(* IEC 61131-3 sources: daoli-st-library/DL_Process (part 32) *)

(* ---- FB_DL_ElectrolyzerStackPurgeSeq.st ---- *)
//==============================================================================
// 功能块：FB_DL_ElectrolyzerStackPurgeSeq ｜ 中文名称：电解槽氮气吹扫与升压序（复杂度 C4）
// 所属子库：DL_Process ｜ 版本 VERSION: v1.0.0 ｜ 兼容：CODESYS V3.5+ / TwinCAT 3 / 汇川 InoProShop
// 功能描述：电解槽停机检修后的投运前置序——低压氮气保压检漏 → N2 置换吹扫（按置换
//           倍数 n = ln(C0/C1) 算所需体积）→ O2 校验 → 升压至运行压力 → 就绪放行
//           （H2 侧仅在就绪相且 O2 合格时才允许打开）→ 泄压走 eVent 单向。泄漏率超
//           限、吹扫/升压超时、O2 不合格一律不放行并锁存故障。
// 开源溯源 (Origin)：道莅原创实现（参考 ISO 22734 水电解制氢系统与 GB/T 19774 水
//           电解制氢系统技术要求 分类与参数域，许可证=MIT，借鉴点=「惰性气体置换至
//           爆炸下限以下再投氢」的置换倍数判据与硬互锁序）
// 单位表：O2[%] / 压力[bar] / 流量[Nm³/h] / 体积[Nm³] / 泄漏率[bar/min] / 时间[ms]
// 置换倍数公式（本件核心判据，单位与推导写清）：
//   n = ln(C0 / C1)；C0 = 空气 O2 体积分数 20.9 [%]，C1 = 目标 O2 阈值 1.0 [%]
//   → n = ln(20.9 / 1.0) ≈ 3.04 [倍]，即需通入约 3.04 倍栈容积的 N2。
//   累计 N2 体积 [Nm³] = Σ (fN2FlowNm3h ÷ 3600 × Δt[s])，Δt 取 DL_ELZ_DT_S 假定任务
//   周期 10 ms；置换倍数出口 = 累计体积 ÷ 栈容积 [倍]。除零由段 3/段 4 双侧闸拦。
// 错误码表（Process 段 0005，故障窗口 3F01~3F09，信息窗口 3F81/3F82）：
//   16#0005_3F01 故障级：组态非法（栈容积/目标压/泄漏限/时间量 <= 0 或 O2 阈值域外）
//   16#0005_3F02 故障级：实时量入口非有限（O2 / 压力 / 流量 NaN 或 Inf），拒算
//   16#0005_3F03 故障级：检修保压检漏超限（泄漏率 > fLeakLimitBarPerMin，不放行）
//   16#0005_3F04 故障级：吹扫超时（tPurgeMaxTime 内置换倍数未达 n）
//   16#0005_3F05 故障级：O2 校验失败（校验窗内 O2 未降至阈值以下）
//   16#0005_3F06 故障级：升压超时（预充压或正式升压未达目标压）
//   16#0005_3F07 故障级：投运前保压检漏超限（就绪相保压窗内泄漏率超限，不放行）
//   16#0005_3F08 故障级兜底：状态机落 ELSE 非法态，全输出断
//   16#0005_3F09 故障级：H2 硬互锁违反（就绪相 O2 回升超阈值，立即关 H2 并锁存）
//   16#0005_3F81 信息级：置换倍数达标（置换完成拍，不置 bError）
//   16#0005_3F82 信息级：系统就绪放行（进入 eReady 拍，不置 bError）
//           故障级码全部锁存回放（R187），唯一清除路径 = bReset 上升沿。
// 状态机：E_DL_ElyzPurgeState（八态：eIdle=0 / eLeakTest=10 / ePurge=20 / eVerifyO2=30 /
//           ePressurize=40 / eReady=50 / eVent=60 / eFault=99）。eVent 为单向泄压相，
//           迁出唯一目标 = eIdle，不得返回 eReady（防止带氢泄压后直接投运）。
// 边界行为：① H2 侧硬互锁三重闸：相位必须是 eReady、O2 <= 阈值、无任何故障锁存；段 8
//           的 CASE ELSE 与出口断言各断一次（双保险）；② O2 未达标绝不进 eReady，故
//           不可能放 H2；③ 泄漏率判据只用「>」单侧直比（泄漏率本身是统计量，不设容差
//           死区，避免漏判）；④ 八态 CASE 每态显式 + ELSE 兜底 → 3F08 全断；⑤ 中止在
//           任何运行相都只迁入 eVent（单向泄压），不走「原地停机」路径。
// 语义假设：① fO2Pct 为栈内气相 O2 体积分数，单位 %；② fLeakDropBarPerMin 由上层
//           压降速率仪表或本库泄漏率估算件提供（本件不重复实现估算）；③ N2 流量为
//           标况体积流量，压力对体积的修正由上层完成；④ 栈容积含管路死体积。
// 依赖纪律：仅 Standard.library（TON / R_TRIG / LN）；零 GVL、零 VAR_EXTERNAL、零物
//           理地址直连，业务侧只经引脚注入。
// 修订历史：v1.0.0 2026-11-25 R88 首版（无人值守批次 · 复杂件 C4 · 序号 3）
//==============================================================================

(*------------------------------------------------------------------------------
 * 枚举: E_DL_ElyzPurgeState（归属本功能块，同文件发布，全库唯一定义）
 * 含义: 吹扫升压相位，与段 7 状态机、段 8 输出置位一一对应。
 *-----------------------------------------------------------------------------*)
TYPE E_DL_ElyzPurgeState :
(
    eIdle       := 0,  // 空闲：等启动沿 / Idle, awaiting the start edge
    eLeakTest   := 10, // 检修检漏：低压氮气保压测泄漏率 / Leak test at low nitrogen pressure
    ePurge      := 20, // 吹扫：N2 置换至置换倍数达标 / Purge until the exchange ratio is reached
    eVerifyO2   := 30, // O2 校验：静置取样，O2 须稳定在阈值下 / O2 verification with a stable sample
    ePressurize := 40, // 升压：N2 升至运行压力 / Pressurise to the operating pressure
    eReady      := 50, // 就绪：放行相，H2 侧唯一允许投运的相位 / Ready, the only phase allowing H2
    eVent       := 60, // 泄压：单向排空至常压 / Vent, one-way depressurisation
    eFault      := 99  // 故障：泄漏/超时/O2/互锁/非法态 / Fault, leak, timeout, O2, interlock or illegal state
);
END_TYPE

FUNCTION_BLOCK FB_DL_ElectrolyzerStackPurgeSeq
VAR_INPUT
    xEnable             : BOOL;   // 使能，FALSE 期间按中止处理（转泄压） [—] / Enable, a drop aborts into venting
    xStart              : BOOL;   // 启动请求，上升沿生效 [—] / Start request, rising edge effective
    xAbort              : BOOL;   // 中止请求，任意拍生效，转 eVent 单向泄压 [—] / Abort request, moves to one-way venting
    xReset              : BOOL;   // 故障复位，上升沿清全部锁存 [—] / Fault reset, rising edge clears all latches
    fO2Pct              : LREAL;  // 栈内气相 O2 体积分数 [%] / Gas-phase O2 volume fraction [%]
    fStackPressBar      : LREAL;  // 栈内实际压力 [bar] / Actual stack pressure [bar]
    fTargetPressBar     : LREAL;  // 运行目标压力 [bar]，须 > 0 / Operating target pressure [bar]
    fN2FlowNm3h         : LREAL;  // 氮气标况流量 [Nm³/h] / Nitrogen normal-volume flow [Nm3/h]
    fStackVolM3         : LREAL;  // 栈与管路总容积 [Nm³]，须 > 0 / Total stack and piping volume [Nm3]
    fLeakDropBarPerMin  : LREAL;  // 实测压力下降速率 [bar/min] / Measured pressure decay rate [bar/min]
    fLeakLimitBarPerMin : LREAL;  // 允许泄漏率上限 [bar/min]，须 > 0 / Allowed leak rate ceiling [bar/min]
    tPurgeMaxTime       : TIME;   // 吹扫最长允许时间 [ms] / Maximum purge time [ms]
    tHoldTime           : TIME;   // 保压/取样稳定窗 [ms] / Hold and sampling window [ms]
    tPressTimeout       : TIME;   // 升压与预充压超时 [ms] / Pressurisation timeout [ms]
END_VAR
VAR_OUTPUT
    xN2ValveCmd         : BOOL;   // 氮气进气阀命令 [—] / Nitrogen inlet valve command
    xVentValveCmd       : BOOL;   // 排放阀命令（吹扫出口与泄压共用） [—] / Vent valve command
    xH2ValveCmd         : BOOL;   // 氢气侧阀命令（仅就绪相且 O2 合格才允许） [—] / H2 valve, ready phase and O2 proven only
    bRunning            : BOOL;   // 顺控运行中（非空闲非就绪非故障非泄压） [—] / Sequencing active
    bDone               : BOOL;   // 就绪放行电平（eReady 相） [—] / Ready-released level in the eReady phase
    bError              : BOOL;   // 故障级标志，仅故障级码置位 [—] / Fault-class flag, fault-level codes only
    nErrCode            : UDINT;  // 错误码，0 = 无错 [—] / Error code, 0 = none
    fPurgeVolRatio      : LREAL;  // 置换倍数出口 [倍] = 累计 N2 体积 ÷ 栈容积 / Exchange ratio [ratio]
    nPurgeCount         : UDINT;  // 累计吹扫次数 [次] / Accumulated purge count
END_VAR
VAR
    _eState             : E_DL_ElyzPurgeState := E_DL_ElyzPurgeState.eIdle; // 当前相位 [—] / Current phase
    _bInit              : BOOL := FALSE; // 首扫标志，取非判定 [—] / First-scan flag, tested negated
    _fPurgeVolNm3       : LREAL;         // 累计通入氮气体积 [Nm³] / Accumulated nitrogen volume [Nm3]
    _fReqRatioN         : LREAL;         // 所需置换倍数 n = ln(C0/C1) [倍] / Required exchange ratio n [ratio]
    _fPurgeVolRatio     : LREAL;         // 本拍置换倍数 [倍] / Exchange ratio of this scan [ratio]
    _nPurgeCount        : UDINT;         // 内部累计吹扫次数 [次] / Internal purge counter
    _bCfgBad            : BOOL;          // 组态非法锁存 / Illegal configuration latch
    _bCfgOk             : BOOL;          // 本拍组态合法（派生量不锁存） [—] / Configuration legal this scan, derived
    _bSigBad            : BOOL;          // 实时量非有限锁存 / Non-finite process value latch
    _bLeakErr           : BOOL;          // 检修检漏超限锁存 / Commissioning leak-test latch
    _bPurgeTmo          : BOOL;          // 吹扫超时锁存 / Purge timeout latch
    _bO2Err             : BOOL;          // O2 校验失败锁存 / O2 verification failure latch
    _bPressTmo          : BOOL;          // 升压超时锁存 / Pressurisation timeout latch
    _bLeakReadyErr      : BOOL;          // 投运前检漏超限锁存 / Pre-start leak-test latch
    _bH2LockErr         : BOOL;          // H2 互锁违反锁存 / H2 interlock violation latch
    _bIllegal           : BOOL;          // 非法状态标志 / Illegal state flag
    _bInfoRatio         : BOOL;          // 置换达标信息当拍标志 / Ratio-reached info flag of this scan
    _bInfoReady         : BOOL;          // 就绪放行信息当拍标志 / Ready info flag of this scan
    _bAbortReq          : BOOL;          // 中止请求合成（xAbort 或失能） [—] / Combined abort request
    _bO2Ok              : BOOL;          // O2 合格判据（派生量） [—] / O2 proven criterion, derived
    _bH2Permit          : BOOL;          // H2 投运许可（三重闸合成） [—] / H2 permit, three gates combined
    rtStart             : R_TRIG;        // 启动沿，段 6 无条件刷新 [—] / Start edge, refreshed in segment 6
    rtReset             : R_TRIG;        // 复位沿，段 6 无条件刷新 [—] / Reset edge, refreshed in segment 6
    tonLeakFill         : TON;           // 检修预充压超时 [ms] / Commissioning pre-fill timeout [ms]
    tonHold             : TON;           // 检修保压窗 [ms] / Commissioning hold window [ms]
    tonPurgeMax         : TON;           // 吹扫最长允许时间 [ms] / Maximum purge time [ms]
    tonO2Win            : TON;           // O2 合格稳定窗 [ms] / O2 stability window [ms]
    tonO2Max            : TON;           // O2 校验最长等待 [ms] / Maximum O2 verification wait [ms]
    tonPress            : TON;           // 升压超时 [ms] / Pressurisation timeout [ms]
    tonReadyHold        : TON;           // 就绪相保压窗 [ms] / Ready-phase hold window [ms]
END_VAR
VAR CONSTANT
    DL_EPS                : LREAL := 1.0E-9;  // 浮点容差零点，兼作除法分母下限 / Float epsilon, also the divisor floor
    DL_ELZ_O2_AIR_PCT     : LREAL := 20.9;    // 空气 O2 体积分数 C0 [%] / O2 fraction of air C0 [%]
    DL_ELZ_O2_LIMIT_PCT   : LREAL := 1.0;     // 投运前 O2 阈值 C1 [%] / O2 limit before start-up C1 [%]
    DL_ELZ_SEC_PER_H      : LREAL := 3600.0;  // 小时折算秒 [s/h]，流量积分用 / Seconds per hour for the flow integral
    DL_ELZ_DT_S           : LREAL := 0.01;    // 体积积分假定任务周期 [s]（10 ms） / Assumed task period for the volume integral [s]
    DL_ELZ_LEAK_PRESS_BAR : LREAL := 2.0;     // 检修检漏预充压 [bar] / Commissioning leak-test pressure [bar]
    DL_ELZ_PRESS_TOL_BAR  : LREAL := 0.5;     // 升压到位容差 [bar] / Pressurisation tolerance [bar]
    DL_ELZ_VENT_DONE_BAR  : LREAL := 0.20;    // 泄压完成阈值 [bar] / Vent completion threshold [bar]
    DL_ELZ_PRESS_MAX_BAR  : LREAL := 400.0;   // 压力反馈合法幅值上限 [bar] / Legal pressure ceiling [bar]
END_VAR

(*------------------------------------------------------------------------------
 * 段 1｜每拍预置：全部输出先落安全侧（H2 阀优先断），单拍标志预清零
 *      All outputs preset to the safe side, the H2 valve first, one-shot flags cleared
 *-----------------------------------------------------------------------------*)
xH2ValveCmd := FALSE;                       // 氢气阀先断（最高优先级安全侧） / H2 valve cleared first
xN2ValveCmd := FALSE; xVentValveCmd := FALSE; // 氮气与排放阀先断 / Nitrogen and vent valves cleared
bRunning := FALSE;  bDone := FALSE;         // 运行与就绪标志每拍重算 / Running and ready flags recomputed
bError := FALSE;    nErrCode := 16#0000_0000; // 故障标志与错误码每拍重算 / Fault flag and code recomputed
_bIllegal := FALSE; _bInfoRatio := FALSE; _bInfoReady := FALSE; // 非法态与两条信息标志预清零 / Illegal and info flags pre-cleared

(*------------------------------------------------------------------------------
 * 段 2｜首扫初始化：所需置换倍数 n = ln(C0/C1) 只算一次，计数与体积清零
 *      First-scan initialisation, the required ratio n computed once
 *-----------------------------------------------------------------------------*)
IF NOT _bInit THEN
    _eState     := E_DL_ElyzPurgeState.eIdle; // 相位从空闲起步 / Phase starts idle
    _fPurgeVolNm3 := 0.0;  _nPurgeCount := 0; // 累计体积与吹扫次数清零 / Volume and purge counter at zero
    _fReqRatioN := 0.0;                       // 置换倍数先清零 / Required ratio starts at zero
    IF DL_ELZ_O2_LIMIT_PCT > DL_EPS THEN
        _fReqRatioN := LN(DL_ELZ_O2_AIR_PCT / DL_ELZ_O2_LIMIT_PCT); // n = ln(C0/C1) ≈ 3.04 [倍]，除数已判零 / Ratio n, divisor already proven
    END_IF
    _bInit := TRUE;                           // 首扫只做一次 / The first scan runs once
END_IF

(*------------------------------------------------------------------------------
 * 段 3｜实时量入口非有限闸 + 组态闸（O2 阈值域闸与除零闸并列）
 *      Non-finite inlet gate and configuration gates
 *-----------------------------------------------------------------------------*)
IF NOT (fO2Pct > -1.0E30 AND fO2Pct < 1.0E30) THEN _bSigBad := TRUE; END_IF            // O2 非有限 → 3F02 / Non-finite O2, 3F02
IF NOT (fStackPressBar > -1.0E30 AND fStackPressBar < 1.0E30) THEN _bSigBad := TRUE; END_IF // 压力非有限 → 3F02 / Non-finite pressure, 3F02
IF ABS(fStackPressBar) > DL_ELZ_PRESS_MAX_BAR THEN _bSigBad := TRUE; END_IF             // 压力幅值超上限 → 3F02 / Beyond the ceiling, 3F02
IF NOT (fN2FlowNm3h > -1.0E30 AND fN2FlowNm3h < 1.0E30) OR (fN2FlowNm3h < 0.0) THEN _bSigBad := TRUE; END_IF // 流量非有限或负值 → 3F02 / Non-finite or negative flow, 3F02
IF NOT (fStackVolM3 > -1.0E30 AND fStackVolM3 < 1.0E30) THEN _bCfgBad := TRUE; END_IF   // 栈容积非有限 → 3F01 / Non-finite volume, 3F01
IF NOT (fTargetPressBar > -1.0E30 AND fTargetPressBar < 1.0E30) THEN _bCfgBad := TRUE; END_IF // 目标压非有限 → 3F01 / Non-finite target, 3F01
IF (fStackVolM3 <= DL_EPS) OR (fTargetPressBar <= DL_EPS) OR (fLeakLimitBarPerMin <= DL_EPS) THEN _bCfgBad := TRUE; END_IF // 三者须为正 → 3F01 / All three must be positive
IF NOT (fLeakDropBarPerMin > -1.0E30 AND fLeakDropBarPerMin < 1.0E30) THEN _bSigBad := TRUE; END_IF // 泄漏率非有限 → 3F02（R88 修复：原漏项致 NaN 判合格） / non-finite leak rate, 3F02
IF (fO2Pct < 0.0) OR (fO2Pct > 100.0) THEN _bSigBad := TRUE; END_IF                    // O2 超出 0~100% 域 → 3F02 / O2 outside 0..100, 3F02
IF (tPurgeMaxTime <= T#0MS) OR (tHoldTime <= T#0MS) OR (tPressTimeout <= T#0MS) THEN _bCfgBad := TRUE; END_IF // 时间量须为正 → 3F01 / Time values must be positive
_bCfgOk := NOT _bCfgBad;                    // 本拍组态合法派生量 / Configuration-legal derived flag of this scan
_bO2Ok  := (fO2Pct <= DL_ELZ_O2_LIMIT_PCT) AND (NOT _bSigBad); // O2 合格判据（非有限时不判合格） / O2 proven unless non-finite

(*------------------------------------------------------------------------------
 * 段 4｜吹扫体积积分与置换倍数（除零双侧闸：栈容积与秒折算均先判分母）
 *      Purge volume integral and the exchange ratio, both divisors proven first
 *-----------------------------------------------------------------------------*)
IF (_eState = E_DL_ElyzPurgeState.ePurge) AND (NOT _bCfgBad) THEN
    IF DL_ELZ_SEC_PER_H > DL_EPS THEN
        _fPurgeVolNm3 := _fPurgeVolNm3 + (fN2FlowNm3h / DL_ELZ_SEC_PER_H) * DL_ELZ_DT_S; // 体积积分 [Nm³] / Volume integral [Nm3]
    END_IF
END_IF
_fPurgeVolRatio := 0.0;                     // 置换倍数先清零 / Exchange ratio pre-cleared
IF fStackVolM3 > DL_EPS THEN
    _fPurgeVolRatio := _fPurgeVolNm3 / fStackVolM3; // 置换倍数 [倍] = 累计体积 ÷ 栈容积 / Ratio = volume over stack volume
END_IF
fPurgeVolRatio := _fPurgeVolRatio;          // 置换倍数出口 [倍] / Exchange ratio outlet [ratio]

(*------------------------------------------------------------------------------
 * 段 5｜中止入口（任意运行相 → eVent 单向泄压）与复位
 *      Abort entry into one-way venting plus the reset edge
 *-----------------------------------------------------------------------------*)
_bAbortReq := xAbort OR (NOT xEnable);      // 中止请求合成：显式中止或失能 / Combined abort: explicit abort or enable loss
IF _bAbortReq AND (_eState <> E_DL_ElyzPurgeState.eIdle)
   AND (_eState <> E_DL_ElyzPurgeState.eVent) AND (_eState <> E_DL_ElyzPurgeState.eFault) THEN
    _eState := E_DL_ElyzPurgeState.eVent;   // 转单向泄压相（禁原地停机） / Move to one-way venting, never a plain stop
END_IF
IF rtReset.Q THEN
    _bCfgBad := FALSE;  _bSigBad := FALSE;  _bLeakErr := FALSE; // 复位清组态/入口/检漏锁存 / Clears configuration, inlet and leak latches
    _bPurgeTmo := FALSE; _bO2Err := FALSE; _bPressTmo := FALSE;  // 复位清吹扫/校验/升压锁存 / Clears purge, O2 and pressure latches
    _bLeakReadyErr := FALSE; _bH2LockErr := FALSE;               // 复位清投运检漏与互锁锁存 / Clears pre-start leak and interlock latches
END_IF

(*------------------------------------------------------------------------------
 * 段 6｜定时器与边沿无条件周期刷新（R7：CASE 之外每拍必调，各司其职不复用）
 *      Timers and edges refreshed unconditionally every scan, outside the CASE
 *-----------------------------------------------------------------------------*)
rtStart(CLK := xStart); rtReset(CLK := xReset); // 启动沿与复位沿无条件刷新 / Start and reset edges refreshed
tonLeakFill(IN := (_eState = E_DL_ElyzPurgeState.eLeakTest) AND (fStackPressBar < DL_ELZ_LEAK_PRESS_BAR), PT := tPressTimeout); // 检修预充压超时
tonHold(IN := (_eState = E_DL_ElyzPurgeState.eLeakTest) AND (fStackPressBar >= DL_ELZ_LEAK_PRESS_BAR), PT := tHoldTime);       // 检修保压窗
tonPurgeMax(IN := (_eState = E_DL_ElyzPurgeState.ePurge), PT := tPurgeMaxTime);   // 吹扫最长允许时间 / Maximum purge time
tonO2Win(IN := (_eState = E_DL_ElyzPurgeState.eVerifyO2) AND _bO2Ok, PT := tHoldTime); // O2 合格稳定窗 / O2 stability window
tonO2Max(IN := (_eState = E_DL_ElyzPurgeState.eVerifyO2), PT := tPurgeMaxTime);       // O2 校验最长等待 / Maximum O2 wait
tonPress(IN := (_eState = E_DL_ElyzPurgeState.ePressurize), PT := tPressTimeout);     // 升压超时 / Pressurisation timeout
tonReadyHold(IN := (_eState = E_DL_ElyzPurgeState.eReady), PT := tHoldTime);          // 就绪相保压窗 / Ready hold window

(*------------------------------------------------------------------------------
 * 段 7｜状态机（每态显式迁移判据，ELSE 兜底落故障）
 *      Phase machine with explicit transition criteria and an ELSE fallback
 *-----------------------------------------------------------------------------*)
CASE _eState OF
    E_DL_ElyzPurgeState.eIdle:              // 空闲：启动沿 + 组态合法 + 入口可用才进检漏 / Idle, legal start edge only
        IF rtStart.Q AND _bCfgOk AND (NOT _bSigBad) AND (NOT _bAbortReq) THEN
            _fPurgeVolNm3 := 0.0;           // 新循环体积清零 / Volume reset for the new cycle
            _eState := E_DL_ElyzPurgeState.eLeakTest; // 进检修检漏相 / To the leak-test phase
        END_IF
    E_DL_ElyzPurgeState.eLeakTest:          // 检修检漏：保压窗满判泄漏率，超限不放行 / Leak rate judged at the end of the hold
        IF (fStackPressBar < DL_ELZ_LEAK_PRESS_BAR) AND tonLeakFill.Q THEN
            _bPressTmo := TRUE; _eState := E_DL_ElyzPurgeState.eFault; // 预充压超时 → 3F06 / Pre-fill timeout, 3F06
        ELSIF tonHold.Q THEN
            IF NOT (fLeakDropBarPerMin <= fLeakLimitBarPerMin) THEN // fail-closed：非有限时 NOT(FALSE)=TRUE 即判超限（R88 修复）
                _bLeakErr := TRUE; _eState := E_DL_ElyzPurgeState.eFault; // 泄漏率超限 → 3F03 / Leak over limit, 3F03
            ELSE
                _eState := E_DL_ElyzPurgeState.ePurge; // 检漏合格，进吹扫相 / Leak proven, to purge
            END_IF
        END_IF
    E_DL_ElyzPurgeState.ePurge:             // 吹扫：置换倍数达 n 即完成，超时落故障 / Purge until the ratio reaches n
        IF _fPurgeVolRatio >= _fReqRatioN THEN
            _nPurgeCount := _nPurgeCount + 1;  // 吹扫次数递增 / Purge counter incremented
            _bInfoRatio  := TRUE;              // 置换达标信息 / Ratio-reached info
            _eState      := E_DL_ElyzPurgeState.eVerifyO2; // 进 O2 校验相 / To O2 verification
        ELSIF tonPurgeMax.Q THEN
            _bPurgeTmo := TRUE; _eState := E_DL_ElyzPurgeState.eFault; // 吹扫超时 → 3F04 / Purge timeout, 3F04
        END_IF
    E_DL_ElyzPurgeState.eVerifyO2:          // O2 校验：稳定窗满即合格，最长等待到则失败 / Stable window or maximum wait
        IF tonO2Win.Q THEN
            _eState := E_DL_ElyzPurgeState.ePressurize; // O2 合格稳定，进升压相 / O2 proven, to pressurise
        ELSIF tonO2Max.Q THEN
            _bO2Err := TRUE; _eState := E_DL_ElyzPurgeState.eFault; // 校验失败 → 3F05 / Verification failed, 3F05
        END_IF
    E_DL_ElyzPurgeState.ePressurize:        // 升压：达目标压容差即就绪，超时落故障 / Pressurise to the target band
        IF fStackPressBar >= (fTargetPressBar - DL_ELZ_PRESS_TOL_BAR) THEN
            _bInfoReady := TRUE;            // 就绪放行信息 / Ready info
            _eState     := E_DL_ElyzPurgeState.eReady; // 进就绪相 / To the ready phase
        ELSIF tonPress.Q THEN
            _bPressTmo := TRUE; _eState := E_DL_ElyzPurgeState.eFault; // 升压超时 → 3F06 / Pressurisation timeout, 3F06
        END_IF
    E_DL_ElyzPurgeState.eReady:             // 就绪：O2 回升即互锁故障；保压窗满判泄漏；启动撤销回空闲
        IF NOT _bO2Ok THEN
            _bH2LockErr := TRUE; _eState := E_DL_ElyzPurgeState.eFault; // O2 回升，H2 互锁违反 → 3F09 / O2回升, 3F09
        ELSIF tonReadyHold.Q AND (NOT (fLeakDropBarPerMin <= fLeakLimitBarPerMin)) THEN // fail-closed 同判据（R88 修复）
            _bLeakReadyErr := TRUE; _eState := E_DL_ElyzPurgeState.eFault; // 投运前检漏超限 → 3F07 / Pre-start leak, 3F07
        ELSIF tonReadyHold.Q AND (NOT xStart) THEN
            _eState := E_DL_ElyzPurgeState.eIdle; // 就绪撤销且检漏合格，回空闲 / Ready withdrawn and leak proven, idle
        END_IF
    E_DL_ElyzPurgeState.eVent:              // 泄压：单向排空至阈值以下才回空闲 / Vent one-way, idle below the threshold
        IF fStackPressBar <= DL_ELZ_VENT_DONE_BAR THEN _eState := E_DL_ElyzPurgeState.eIdle; END_IF
    E_DL_ElyzPurgeState.eFault:             // 故障：复位沿且组态合法且入口可用才回空闲 / Fault, reset edge only
        IF rtReset.Q AND _bCfgOk AND (NOT _bSigBad) THEN _eState := E_DL_ElyzPurgeState.eIdle; END_IF
    ELSE                                    // 非法状态兜底（R6：CASE 必带 ELSE）/ Illegal-state fallback
        _bIllegal := TRUE; _eState := E_DL_ElyzPurgeState.eFault; // 非法态 → 3F08，落故障 / Illegal state, 3F08
END_CASE

(*------------------------------------------------------------------------------
 * 段 8｜输出置位（H2 侧三重闸 + 出口断言双保险；泄压相只开排放阀）
 *      Output assignment, H2 gated threefold with a second outlet assertion
 *-----------------------------------------------------------------------------*)
_bH2Permit := (_eState = E_DL_ElyzPurgeState.eReady) AND _bO2Ok AND (NOT _bAbortReq)
              AND (NOT _bH2LockErr) AND (NOT _bLeakReadyErr); // H2 许可三重闸：相位 + O2 + 无故障 / Three gates: phase, O2, no fault
CASE _eState OF
    E_DL_ElyzPurgeState.eLeakTest:          // 检修检漏：未达预充压才开 N2，排放阀关 / Fill nitrogen until the test pressure
        xN2ValveCmd := (fStackPressBar < DL_ELZ_LEAK_PRESS_BAR); // 达压即关氮气 / Nitrogen closed once at pressure
    E_DL_ElyzPurgeState.ePurge:             // 吹扫：氮气进、排放出，双向流路 / Purge with both inlet and vent open
        xN2ValveCmd := TRUE; xVentValveCmd := TRUE; // 进气与排放同开 / Inlet and vent both open
    E_DL_ElyzPurgeState.eVerifyO2:          // O2 校验：静置取样，两阀均关 / Verification with both valves closed
        xN2ValveCmd := FALSE; xVentValveCmd := FALSE; // 静态取样 / Static sampling
    E_DL_ElyzPurgeState.ePressurize:        // 升压：只开氮气，排放阀必须关 / Pressurise with the vent closed
        xN2ValveCmd := TRUE; xVentValveCmd := FALSE; // 关排放防漏压 / Vent closed to hold pressure
    E_DL_ElyzPurgeState.eReady:             // 就绪：只允许 H2（严格由三重闸决定） / Ready, H2 by the three gates only
        xH2ValveCmd := _bH2Permit;          // H2 阀由许可位驱动 / H2 valve driven by the permit
    E_DL_ElyzPurgeState.eVent:              // 泄压：只开排放阀，N2 与 H2 全关 / Vent only, nitrogen and H2 closed
        xVentValveCmd := TRUE;
    ELSE                                    // 其余相（空闲/故障）全断 / Other phases, all off
        xN2ValveCmd := FALSE; xVentValveCmd := FALSE; xH2ValveCmd := FALSE; // 全阀断 / All valves off
END_CASE
IF NOT _bH2Permit THEN
    xH2ValveCmd := FALSE;                   // 出口断言：许可不成立时 H2 必须为 FALSE / Outlet assertion, H2 false without a permit
END_IF
bRunning := (_eState <> E_DL_ElyzPurgeState.eIdle) AND (_eState <> E_DL_ElyzPurgeState.eReady)
            AND (_eState <> E_DL_ElyzPurgeState.eVent) AND (_eState <> E_DL_ElyzPurgeState.eFault); // 运行标志
bDone := (_eState = E_DL_ElyzPurgeState.eReady); nPurgeCount := _nPurgeCount; // 就绪放行电平与吹扫次数出口 / Ready level and purge count

(*------------------------------------------------------------------------------
 * 段 9｜错误码映射（锁存回放，R187：故障相不按当下输入重推断）
 *      Error-code map, latched replay
 *-----------------------------------------------------------------------------*)
IF _bIllegal THEN nErrCode := 16#0005_3F08; bError := TRUE;        // 故障级兜底：非法态 / Fault, illegal state fallback
ELSIF _bCfgBad THEN nErrCode := 16#0005_3F01; bError := TRUE;      // 故障级：组态非法 / Fault, illegal configuration
ELSIF _bSigBad THEN nErrCode := 16#0005_3F02; bError := TRUE;      // 故障级：入口非有限 / Fault, non-finite inlet
ELSIF _bH2LockErr THEN nErrCode := 16#0005_3F09; bError := TRUE;   // 故障级：H2 硬互锁违反 / Fault, H2 interlock violated
ELSIF _bLeakErr THEN nErrCode := 16#0005_3F03; bError := TRUE;     // 故障级：检修检漏超限 / Fault, commissioning leak
ELSIF _bLeakReadyErr THEN nErrCode := 16#0005_3F07; bError := TRUE; // 故障级：投运前检漏超限 / Fault, pre-start leak
ELSIF _bPurgeTmo THEN nErrCode := 16#0005_3F04; bError := TRUE;    // 故障级：吹扫超时 / Fault, purge timeout
ELSIF _bO2Err THEN nErrCode := 16#0005_3F05; bError := TRUE;       // 故障级：O2 校验失败 / Fault, O2 verification failed
ELSIF _bPressTmo THEN nErrCode := 16#0005_3F06; bError := TRUE;    // 故障级：升压超时 / Fault, pressurisation timeout
ELSIF _bInfoRatio THEN nErrCode := 16#0005_3F81;                   // 信息级：置换倍数达标 / Info, exchange ratio reached
ELSIF _bInfoReady THEN nErrCode := 16#0005_3F82;                   // 信息级：系统就绪放行 / Info, ready released
END_IF
END_FUNCTION_BLOCK

(* ---- FB_DL_ElTestStation.st ---- *)
(*
  FB_DL_ElTestStation  —  EL 检测工站（相机触发、缺陷坐标映射、OK/NG 归档） / EL test station: camera trigger, defect coordinate mapping, OK/NG archive
  分类 Category : DL_Process
  版本 Version  : 1.0.1
  来源 Source   : roadmap-pv-p2 — 光伏行业池 EL 检测缺口件
  溯源 Origin   : clean-room 实现，未复制任何源码行
  功能 Function : 1) 五相顺控：eIdle → eTrig（单发相机触发 bCamTrig，等回读
                  bCamDone，tCamTo 超时判）→ eMap（缺陷坐标映射：首缺陷
                  (fDefX,fDefY) 换算单元号 nDefCell，除法前域闸防除零）
                  → eDone（OK/NG 归档出口）→ 回 eIdle；
                  2) NG 判据：uDefCount > 0 且坐标在板面域内 → NG 归档
                  （uNgCount 累计）；uDefCount = 0 → OK 归档（uOkCount 累计）；
                  3) 故障级：0397 触发后超时无回读 / 0398 缺陷坐标越界或
                  非有限锁存（NG 侧防御，归档冻结）/ 0399 组态非法（行列、
                  单元尺寸域）+ ELSE 兜底归并；
                  4) 信息级三码：触发发出 / NG 归档 / OK 归档（单拍沿）；
                  5) 解除式全当拍量（R240 落地），逐 BOOL 标注见段 4。
  边界 Boundary : ① 组态闸：nRows/nCols = 0、fCellW/fCellH <= 0、tCamTo <= 0
                  → 0399 锁存，顺控停发；
                  ② 坐标映射前先做板面域闸（0 <= fDefX < fCellW*nCols 等），
                  域外或非有限 → 0398（NaN 自反判，R79）；TRUNC 前实数域钳制
                  （R151 实数转整数前域钳）；
                  ③ uDefCount 信任来源为相机契约 bCamDone 当拍（头注释声明）；
                  ④ 无 GVL 依赖：纯引脚输入输出，无外部变量引用，无物理 IO 地址。
  依赖 Depends  : Standard.library（TON / R_TRIG）
  码表 Error codes（Process 段 0005，窗口 0397~0399 / 04BF~04C1）:
    16#0005_0397 故障级：触发后超时无回读锁存（tCamTo），锁存至 bReset
    16#0005_0398 故障级：缺陷坐标越界或非有限锁存（防御兜底），锁存至 bReset
    16#0005_0399 故障级：组态非法（行列/单元尺寸/超时域非法）或相位落 ELSE 兜底（归并声明），锁存至 bReset
    16#0005_04BF 信息级：触发发出沿（bCamTrig 单发拍）
    16#0005_04C0 信息级：NG 归档沿（NG 判定拍）
    16#0005_04C1 信息级：OK 归档沿（OK 判定拍）
  修订历史 Revision :
    2026-11-19  v1.0.0  R42 首版（批次 3 · 序号 4）
    2026-11-19  v1.0.1  R42 终审返修：新增段 4A 故障锁存相位迁移闸——0397/0398/0399
                        锁存后 _eState 强制迁 eFault，断 tonCamTo 跨锁存期 IN 保持
                        （否则复位清锁后下一拍 Q 恒 TRUE 立即重锁 0397，解除式不可达），
                        并冻结 eTrig/eMap 相内快照与归档计数副作用；对外引脚契约不变。
*)

TYPE E_DL_EtsState :
(
    eIdle  := 0,     // 空闲：等测试指令 / Idle, waiting test command
    eTrig  := 10,    // 触发：等相机回读 / Trigger, waiting camera readback
    eMap   := 20,    // 映射：缺陷坐标换算单元号 / Map, defect coordinate to cell
    eDone  := 30,    // 完成：归档出口 / Done, archived
    eFault := 90     // 故障：超时或越界锁定 / Fault, latched
);
END_TYPE

FUNCTION_BLOCK FB_DL_ElTestStation
VAR_INPUT
    bTestCmd     : BOOL := FALSE;     // 测试指令，上升沿启动 [-] / Test command edge
    bCamDone     : BOOL := FALSE;     // 相机回读完成（当拍量）[-] / Camera readback done, current-scan
    uDefCount    : UDINT := 0;        // 缺陷点数（bCamDone 当拍采信）[个] / Defect count
    fDefX        : REAL := 0.0;       // 首缺陷 X 坐标 [mm]，板面域 / First defect X coordinate
    fDefY        : REAL := 0.0;       // 首缺陷 Y 坐标 [mm]，板面域 / First defect Y coordinate
    fCellW       : REAL := 50.0;      // 单元宽 [mm]，域 > 0 / Cell width
    fCellH       : REAL := 50.0;      // 单元高 [mm]，域 > 0 / Cell height
    nRows        : USINT := 6;        // 板面单元行数 [个]，域 > 0 / Cell rows
    nCols        : USINT := 10;       // 板面单元列数 [个]，域 > 0 / Cell cols
    tCamTo       : TIME := T#3S;      // 相机回读超时 [ms]，域 > 0 / Camera readback timeout
    bReset       : BOOL := FALSE;     // 复位，上升沿清故障锁存与归档计数 / Reset edge
END_VAR
VAR_OUTPUT
    eState       : E_DL_EtsState;     // 状态出口，段尾单点映射 / State outlet
    bCamTrig     : BOOL;              // 相机触发输出（eTrig 相电平）[-] / Camera trigger output
    nDefCell     : DINT;              // 首缺陷单元号 [0..nRows*nCols-1]，-1 = 无映射 / First defect cell index
    uNgCount     : UDINT;             // NG 归档累计 [片] / NG archive count
    uOkCount     : UDINT;             // OK 归档累计 [片] / OK archive count
    bError       : BOOL;              // 故障锁存标志 / Fault latch flag
    nErrId       : UDINT;             // 事件码，0 = 无事件 / Event code
END_VAR
VAR
    tonCamTo     : TON;               // 相机回读超时（单相独占），无条件刷新 / Camera timeout
    rtTestCmd    : R_TRIG;            // 测试指令沿实例，无条件刷新 / Test command edge instance
    rtReset      : R_TRIG;            // 复位沿实例，无条件刷新 / Reset edge instance
    _eState      : E_DL_EtsState := E_DL_EtsState.eIdle;  // 内部相位（CASE 唯一写入目标）/ Internal phase
    _bTrigSent   : BOOL;              // 触发单发标志（eTrig 相内保持）/ Trigger one-shot flag
    _uDefSnap    : UDINT;             // 缺陷点数采信快照（锁存量）/ Defect count trusted snapshot
    _fXSnap      : REAL;              // 首缺陷 X 采信快照 [mm]（锁存量）/ First defect X snapshot
    _fYSnap      : REAL;              // 首缺陷 Y 采信快照 [mm]（锁存量）/ First defect Y snapshot
    _bNonFin     : BOOL;              // 坐标非有限当拍量 [-] / Non-finite coordinate flag
    _bInPanel    : BOOL;              // 坐标在板面域当拍量 [-] / Coordinate-in-panel flag
    _bFault      : BOOL;              // 故障锁存位（锁存量）/ Latched fault bit
    _uFault      : UDINT;             // 故障码锁存（锁存量）/ Latched fault code
    _uInfo       : UDINT;             // 信息码，每拍重算 / Transient info code
END_VAR

(* —— 段 0：定时器与沿实例无条件周期刷新（禁置于 IF/CASE 内） —— *)
_bNonFin := (fDefX <> fDefX) OR (fDefY <> fDefY)
         OR ((fDefX - fDefX) <> (fDefX - fDefX))
         OR ((fDefY - fDefY) <> (fDefY - fDefY));        // 坐标非有限防御（NaN 自反 + 差值自减）
_bInPanel := (NOT _bNonFin) AND (fDefX >= 0.0) AND (fDefX < fCellW * UDINT_TO_REAL(UINT(nCols)))
          AND (fDefY >= 0.0) AND (fDefY < fCellH * UDINT_TO_REAL(UINT(nRows)));
                                        // 坐标在板面域（当拍量，NaN 与一切比较 FALSE 故先排非有限）
rtTestCmd(CLK := bTestCmd);             // 测试沿（每拍必调）
rtReset(CLK := bReset);                 // 复位沿（每拍必调）
tonCamTo(IN := (_eState = E_DL_EtsState.eTrig), PT := tCamTo);   // 回读超时（单相独占）

(* —— 段 1：单拍量预清零（锁存量 _bFault/_uFault 与采信快照不入清单，禁同拍抹除） —— *)
_uInfo := 16#0000_0000;             // 信息码每拍重算
bCamTrig := FALSE;                  // 触发输出缺省 FALSE（单相承载）
nDefCell := -1;                     // 单元号缺省 -1
nErrId := 16#0000_0000;             // 事件码缺省无事件

(* —— 段 2：复位沿 + 组态域闸（判据当拍量） —— *)
IF rtReset.Q THEN                   // rtReset.Q = 当拍量
    _bFault := FALSE;               // 清故障锁存位
    _uFault := 16#0000_0000;        // 清故障锁存码
    _bTrigSent := FALSE;            // 触发单发标志清零
    uNgCount := 16#0000_0000;       // NG 累计清零
    uOkCount := 16#0000_0000;       // OK 累计清零
END_IF
IF (nRows = 0) OR (nCols = 0) OR (fCellW <= 0.0) OR (fCellH <= 0.0)
   OR (TIME_TO_DINT(tCamTo) <= 0) THEN
    _uFault := 16#0005_0399;        // 故障级：组态非法
    _bFault := TRUE;                // 故障标志与码位配对（R45）
END_IF

(* —— 段 3：回读超时与坐标防御锁存（判据当拍量） —— *)
IF (NOT _bFault) AND tonCamTo.Q THEN
    _uFault := 16#0005_0397;        // 故障级：触发后超时无回读
    _bFault := TRUE;
END_IF
IF (NOT _bFault) AND (_eState = E_DL_EtsState.eMap) AND ((_bNonFin) OR (NOT _bInPanel)) THEN
    _uFault := 16#0005_0398;        // 故障级：坐标越界或非有限
    _bFault := TRUE;
END_IF

(* —— 段 4：故障解除式（R240 落地，逐 BOOL 标注）：
     rtReset.Q = 当拍量；NOT bTestCmd = 当拍量；NOT bCamDone = 当拍量。
     均不含锁存量（_bFault/_uFault），解除边真实可达（指令撤销 + 复位沿）。 —— *)
IF rtReset.Q AND (NOT bTestCmd) AND (NOT bCamDone) THEN
    _bFault := FALSE;               // 清故障锁存位（锁存量，仅此当拍量解除沿可清）
    _uFault := 16#0000_0000;        // 清故障锁存码（锁存量，仅本当拍量解除沿可清）
    IF _eState = E_DL_EtsState.eFault THEN
        _eState := E_DL_EtsState.eIdle;     // 故障相迁出：回空闲
    END_IF
END_IF

(* —— 段 4A：故障锁存相位迁移闸（R42 终审返修，v1.0.1）：
     锁存置位而相位未迁出（0397 超时相 eTrig / 0398 越界相 eMap / 0399 组态任意相）
     时强制入故障相：断 tonCamTo 跨锁存期 IN 保持（IN 恒 TRUE 则 Q 恒 TRUE，
     复位清锁后下一拍立即重锁，解除式不可达），并冻结 eTrig/eMap 相内快照
     与归档副作用；置于段 4 之后，解除沿当拍清锁不触发迁移，无同拍抢迁。 —— *)
IF _bFault AND (_eState <> E_DL_EtsState.eFault) THEN
    _eState := E_DL_EtsState.eFault;        // 锁存即入故障相（锁存量 _bFault 仅解除沿可清，迁移保持至解除）
END_IF

(* —— 段 5：相位机（CASE 全覆盖 + ELSE 兜底） —— *)
CASE _eState OF

E_DL_EtsState.eIdle:
    IF rtTestCmd.Q AND (NOT _bFault) THEN
        _bTrigSent := FALSE;            // 单发标志复位（进相预置）
        _eState := E_DL_EtsState.eTrig; // 进触发相
    END_IF

E_DL_EtsState.eTrig:
    bCamTrig := TRUE;                   // 触发电平（相承载）
    IF NOT _bTrigSent THEN
        _uInfo := 16#0005_04BF;         // 信息级：触发发出沿（进相首拍单发）
        _bTrigSent := TRUE;             // 单发标志
    END_IF
    IF bCamDone THEN                    // 回读完成（当拍量）：采信契约快照
        bCamTrig := FALSE;              // 触发撤销
        _uDefSnap := uDefCount;         // 缺陷数快照（锁存量，仅此处写）
        _fXSnap := fDefX;               // X 快照（锁存量，仅此处写）
        _fYSnap := fDefY;               // Y 快照（锁存量，仅此处写）
        _eState := E_DL_EtsState.eMap;  // 进映射相
    END_IF
    (* 回读超时迁出在段 3 承载 *)

E_DL_EtsState.eMap:
    IF (_bNonFin) OR (NOT _bInPanel) THEN
        ;                               // 越界/非有限迁出在段 3 承载（映射冻结）
    ELSE
        IF _uDefSnap > 0 THEN           // NG 判据（快照域）
            nDefCell := TRUNC(_fXSnap / fCellW) + TRUNC(_fYSnap / fCellH) * USINT_TO_DINT(nCols);
                                        // 单元号映射（域闸已保分母 > 0 与商 < 行列数，无越界；TRUNC 向零取整）
            uNgCount := uNgCount + 1;   // NG 累计递增
            _uInfo := 16#0005_04C0;     // 信息级：NG 归档沿
        ELSE
            uOkCount := uOkCount + 1;   // OK 累计递增
            _uInfo := 16#0005_04C1;     // 信息级：OK 归档沿
        END_IF
        _eState := E_DL_EtsState.eDone; // 进完成相
    END_IF

E_DL_EtsState.eDone:
    IF NOT bTestCmd THEN                // 测试指令撤销：回空闲
        _eState := E_DL_EtsState.eIdle;
    END_IF

E_DL_EtsState.eFault:
    ;                                   // 故障相：归档冻结，等解除沿（段 4 承载迁出）

ELSE
    _uFault := 16#0005_0399;            // 故障级：非法相位兜底（归并组态码，码表声明）
    _bFault := TRUE;
    _eState := E_DL_EtsState.eFault;    // 强制回故障相

END_CASE

(* —— 段 6：出口单点映射（名实同源；锁存码回放，禁同拍抹除） —— *)
IF _bFault THEN
    nErrId := _uFault;              // 故障锁存码回放
    bCamTrig := FALSE;              // 故障相触发输出强制 FALSE（安全侧）
    nDefCell := -1;                 // 故障相单元号恢复哨兵
ELSE
    nErrId := _uInfo;               // 信息码
END_IF
bError := _bFault;                  // 故障标志与锁存位同源
eState := _eState;                  // 状态出口单点映射

END_FUNCTION_BLOCK

(* ---- FB_DL_EmoAndonFab.st ---- *)
// =====================================================================
// FB_DL_EmoAndonFab.st
// 洁净室 EMO-安灯联动呼叫（EMO 急停优先仲裁 + 门审计联动 + 应答/复位管理）
// Cleanroom EMO andon linkage with priority arbitration and door audit
// 所属子库: DL_Process    版本: v1.0.0    兼容: CODESYS V3.5+ / TwinCAT 3 / 汇川 InoProShop
// 码位: 16#0005_047B ~ 16#0005_047F (本件独占 5 槽, 勿复用)
// 溯源: 道莅 clean-room 防御性实现
//       来源组标签: semiconductor, andon, emo, safety-linkage
// 枚举属主: E_DL_AndonLevel —— 全库唯一属主为 DL_Process 安灯呼叫系统件,
//           本件只引用不重声明
// 修改记录: R30 初版 (ROUND_PLAN_R30 序 10)
// 分层声明: 本件为联动编排件, 四级仲裁律全部消费库内安灯呼叫系统件的
//           E_DL_AndonLevel 契约, 不重写普通呼叫仲裁; EMO 触发不唯一属主,
//           首出定位到按钮号; 门审计事件经门开位掩码引脚注入
// =====================================================================
FUNCTION_BLOCK FB_DL_EmoAndonFab
VAR_INPUT
    abEmo        : ARRAY[1..6] OF BOOL;  // EMO 急停按钮阵列 / EMO button array
    bDoorOpenMask: WORD := 0;        // 安全门开位掩码注入, 位 0..5 对应门 1..6 / Door-open mask injected, bit0..5 = door 1..6
    bAck         : BOOL := FALSE;    // 呼叫应答命令 / Call acknowledge command
    bReset       : BOOL := FALSE;    // 事件复位命令 / Event reset command
END_VAR
VAR_OUTPUT
    eAndonLevel  : E_DL_AndonLevel := E_DL_AndonLevel.eNone;  // 联动安灯级别 / Linked andon level
    bLampRed     : BOOL := FALSE;    // 红灯输出 / Red lamp output
    bBuzzer      : BOOL := FALSE;    // 蜂鸣输出（应答后静音）/ Buzzer output, muted after ack
    uFirstEmo    : USINT := 0;       // 首出 EMO 按钮号 1~6, 0 = 无 / First-out EMO button, 0 = none
    eErr         : UDINT := 16#0005_047B;  // 错误码 / Error code
END_VAR
VAR
    rtrAck       : R_TRIG;           // 应答沿检测, 每拍无条件刷新 / Ack edge, refreshed every cycle
    rtrReset     : R_TRIG;           // 复位沿检测, 每拍无条件刷新 / Reset edge, refreshed every cycle
    bEmoAny      : BOOL := FALSE;    // 任一 EMO 有效标记 / Any EMO active flag
    uFirstThis   : USINT := 0;       // 本拍首出候选按钮号 / First-out candidate this cycle
    uFirstLatch  : USINT := 0;       // 首出锁存按钮号 / First-out latched button
    bAckLatch    : BOOL := FALSE;    // 应答静音锁存 / Acknowledge mute latch
    uZi          : INT   := 1;       // 1..6 数组下标 / Array subscript 1..6
END_VAR

// ---------------------------------------------------------------------
// 代码位表（本件独占, 勿复用）:
//   16#0005_047B 信息 无 EMO 无门审计事件
//   16#0005_047C 故障 EMO 急停触发（任一按钮有效, 优先级高于门审计）,
//                解除式 = 全部按钮释放 且 bReset 上升沿
//   16#0005_047D 故障 安全门审计联动（门开掩码非零）, 解除式 = 门掩码归零
//   16#0005_047E 信息 应答沿确认（事件存续期间的应答统计拍,
//                未应答解除不计入应答统计, 沿用安灯呼叫系统语义）
//   16#0005_047F 信息 复位确认（事件已解除后的复位拍, 清应答锁存）
// ---------------------------------------------------------------------

// ---- EMO 首出候选扫描（升序取最小按钮号）/ EMO first-out candidate scan ----
bEmoAny := FALSE;                   // 标记复位 / Reset flag
uFirstThis := 0;                    // 候选清零 / Clear candidate
FOR uZi := 1 TO 6 DO
    IF abEmo[uZi] THEN
        bEmoAny := TRUE;            // 任一按钮有效 / Any button active
        IF uFirstThis = 0 THEN
            uFirstThis := INT_TO_USINT(uZi);    // 升序首出候选 / Ascending first candidate
        END_IF
    END_IF
END_FOR

// ---- 应答与复位沿实例无条件刷新 / Unconditional ack and reset edge refresh ----
rtrAck(CLK := bAck);
rtrReset(CLK := bReset);

// ---- 首出锁存与解除 / First-out latch and release ----
IF (uFirstLatch = 0) AND bEmoAny THEN
    uFirstLatch := uFirstThis;      // 未锁存才仲裁, 同拍取最小按钮号 / Arbitrate only if unlatched, min button
END_IF
IF NOT bEmoAny THEN
    uFirstLatch := 0;               // 全部释放解除首出锁存 / Release when all clear
END_IF
uFirstEmo := uFirstLatch;           // 输出首出按钮号 / Output first-out button

// ---- 应答锁存管理（未应答解除不计入应答统计: 解除拍自动清锁存）
//      Ack latch management, un-acked release clears latch ----
IF rtrAck.Q AND (bEmoAny OR (bDoorOpenMask <> 0)) THEN
    bAckLatch := TRUE;              // 事件存续期间应答生效 / Ack effective while event present
END_IF
IF (NOT bEmoAny) AND (bDoorOpenMask = 0) THEN
    bAckLatch := FALSE;             // 事件消失清应答锁存 / Clear latch on event clear
END_IF

// ---- 联动级别仲裁: EMO 优先于门审计, 同拍取高者 / Level arbitration: EMO over door ----
IF bEmoAny THEN
    eAndonLevel := E_DL_AndonLevel.eMaint;      // EMO 映射最高优先级维修级 / EMO maps to highest level
ELSIF bDoorOpenMask <> 0 THEN
    eAndonLevel := E_DL_AndonLevel.eDevice;     // 门审计映射设备级 / Door audit maps device level
ELSE
    eAndonLevel := E_DL_AndonLevel.eNone;       // 无事件 / No event
END_IF

// ---- 灯与蜂鸣输出（蜂鸣按级别 CASE 判定, 含 ELSE 兜底）/ Lamp and buzzer with CASE fallback ----
bLampRed := bEmoAny OR (bDoorOpenMask <> 0);    // 红灯: 任一事件点亮 / Lamp on any event
CASE eAndonLevel OF
    E_DL_AndonLevel.eNone:     bBuzzer := FALSE;                        // 无事件不鸣响 / No event, silent
    E_DL_AndonLevel.eMaterial: bBuzzer := FALSE;                        // 本件不消费普通缺料级 / Material level not consumed here
    E_DL_AndonLevel.eQuality:  bBuzzer := FALSE;                        // 本件不消费普通品质级 / Quality level not consumed here
    E_DL_AndonLevel.eDevice:   bBuzzer := bLampRed AND (NOT bAckLatch); // 设备级: 未应答鸣响 / Device level: buzzer until ack
    E_DL_AndonLevel.eMaint:    bBuzzer := bLampRed AND (NOT bAckLatch); // 维修级: 未应答鸣响 / Maint level: buzzer until ack
    ELSE                       bBuzzer := bLampRed;                     // 兜底: 未知级别按最响处理 / Fallback: loudest
END_CASE

// ---- 错误码仲裁 / Error arbitration ----
IF bEmoAny THEN
    eErr := 16#0005_047C;           // EMO 触发（最高优先级）/ EMO active, highest priority
ELSIF rtrAck.Q AND bLampRed THEN
    eErr := 16#0005_047E;           // 应答沿确认拍 / Ack edge cycle
ELSIF bDoorOpenMask <> 0 THEN
    eErr := 16#0005_047D;           // 门审计联动 / Door audit linkage
ELSIF rtrReset.Q AND (NOT bEmoAny) THEN
    eErr := 16#0005_047F;           // 复位确认拍 / Reset confirm cycle
ELSE
    eErr := 16#0005_047B;           // 无事件 / No event
END_IF

END_FUNCTION_BLOCK

(* ---- FB_DL_EnergyKpiAggregator.st ---- *)
(*==============================================================================
 * 组件名称 (Component)  : FB_DL_EnergyKpiAggregator
 * 溯源说明 (Provenance) : 道莅 clean-room 防御性实现（PackML 深化）
 * 所属子库 (Sublibrary) : DL_Process / Kpi
 * 当前版本 (Version)    : 1.0.0
 * 兼容性   (Platform)   : CODESYS 3.5 / TwinCAT 3 / 汇川 InoProShop；
 *                         纯 IEC 61131-3（第 3 版），仅用标准库 TON
 * 组件分类 (Category)   : 功能块（FUNCTION_BLOCK）· 单位产量能耗 KPI 聚合
 * 功能一句话 (Summary)  : KPI 窗口内电能累计除以产量计数，得 kWh 每千件。
 * 边界与安全 (Boundary) : ①能量增量小于 0 视为表翻转拒收并置码；
 *                         ②NaN 能量增量拒收（自反判）；
 *                         ③窗口产量为 0 → 保持上次 KPI + 零产量掩码（不做除零）；
 *                         ④KPI 窗口 TON 无条件周期刷新；
 *                         ⑤bReset 清全部窗口累计与有效标志。
 * 错误码    : 16#0005_0365 能量增量非法（负值表翻转或 NaN）——故障级（单拍）
 *             16#0005_0366 零产量掩码激活（窗口产量为 0）——信息级（持续态）
 * 码位总账  : 16#0005_0365 用 / 16#0005_0366 用
 * 修改记录  : v1.0.0 R26 初版
 *==============================================================================*)
FUNCTION_BLOCK FB_DL_EnergyKpiAggregator
VAR_INPUT
    fEnergyDelta : LREAL; // 周期电能增量 [kWh] / Per-cycle energy increment [kWh]
    uProdDelta   : ULINT; // 周期产量增量 [件] / Per-cycle production increment [pcs]
    tKpiWindow   : TIME;  // KPI 统计窗时长 [ms] / KPI window duration [ms]
    bReset       : BOOL;  // 复位：清累计与有效标志 / Reset: clear accumulators and valid flag
END_VAR
VAR_OUTPUT
    fKpi         : LREAL; // 单位产量能耗 [kWh/千件] / Energy per thousand pieces [kWh/kpcs]
    bKpiValid    : BOOL;  // KPI 已有有效结论 / KPI has a valid result
    bZeroProdMask: BOOL;  // 零产量掩码激活 / Zero-production mask active
    eErr         : UDINT; // 本周期错误码，0=无错 / Error code this cycle, 0 = none
END_VAR
VAR
    fEneWin  : LREAL; // 窗内电能累计 [kWh] / In-window energy sum
    uProdWin : ULINT; // 窗内产量累计 [件] / In-window production sum
    tonWin   : TON;   // KPI 窗定时器（无条件刷新）/ KPI window timer
    fEneGrd  : LREAL; // 能量增量守卫副本 / Energy increment guard copy
    fProdReal: LREAL; // 产量实数临时量（除法用）/ Production real temp for division
END_VAR

// ---------- 能量增量防御：负值表翻转与 NaN 拒收 ----------
fEneGrd := fEnergyDelta;
eErr := 0;
IF (fEneGrd <> fEneGrd) OR ((fEneGrd - fEneGrd) <> (fEneGrd - fEneGrd)) THEN
    eErr := 16#0005_0365;                     // NaN 拒收 / NaN rejected
ELSIF fEneGrd < 0.0 THEN
    eErr := 16#0005_0365;                     // 表翻转拒收 / Meter rollover rejected
ELSE
    fEneWin := fEneWin + fEneGrd;             // 合法增量入窗 / Valid increment accumulated
    uProdWin := uProdWin + uProdDelta;        // 产量入窗 / Production accumulated
END_IF

// ---------- 复位：清窗累计与有效标志 ----------
IF bReset THEN
    fEneWin := 0.0;
    uProdWin := ULINT#0;
    fKpi := 0.0;
    bKpiValid := FALSE;
    bZeroProdMask := FALSE;
END_IF

// ---------- 无条件周期刷新：KPI 窗定时器 ----------
tonWin(IN := TRUE, PT := tKpiWindow);

// ---------- 窗到时结算：除法前判零，零产量掩码保持 ----------
IF tonWin.Q THEN
    IF uProdWin > ULINT#0 THEN
        fProdReal := ULINT_TO_LREAL(uProdWin); // 产量实数 / Production as real
        fKpi := fEneWin / (fProdReal / 1000.0); // kWh 每千件（分母前判零）/ kWh per kpcs, zero-guarded
        bKpiValid := TRUE;                    // 有效结论成立 / Valid result set
        bZeroProdMask := FALSE;               // 掩码撤销 / Mask withdrawn
    ELSE
        bZeroProdMask := TRUE;                // 零产量掩码激活 / Zero-production mask
        eErr := 16#0005_0366;                 // 零产量掩码码 / Mask code
        // fKpi 保持上次结论（锁存语义，禁清零）/ fKpi holds last result (no clear)
    END_IF
    fEneWin := 0.0;                           // 窗累计清零 / Window sums cleared
    uProdWin := ULINT#0;
END_IF

END_FUNCTION_BLOCK

(* ---- FB_DL_EnergyMonthPreset.st ---- *)
(*
  ==================================================================
  组件名 Component  : FB_DL_EnergyMonthPreset
  分类   Category   : DL_Process
  版本   Version    : 1.0.0
  功能   Purpose    : 月度能耗预算预置计数与超限预警。月度能耗预算按 12 个月预置表
                      取值（跨月沿自动换表并清零当月累计），能耗增量按脉冲沿累加，
                      出口给出已用 / 剩余 / 占用百分比 / 日均 / 月末预测，并按
                      预警阈与临界阈分四级（正常 / 预警 / 临界 / 超限）。
  溯源   Origin     : 月度预算预置 + 分级预警为本库通用能耗管理语义；本件为
                      clean-room 实现，仅借鉴来源分类与参数域组织（来源标签
                      roadmap-p2-energy），道莅原创设计，未复制任何闭源代码行。
  平台   Platform   : 纯 IEC 61131-3（R_TRIG / REAL 运算，无私有库、无方言转换）
  作者   Author     : 道莅代码库 · PLC 编程专家（R55）
  ------------------------------------------------------------------
  边界 Boundary     :
                      一 本件只做预算计数与分级，不控制用能设备、不发停机命令；
                      二 能耗增量只在 bEnergyPulse 上升沿计入一次（防同拍重复计）；
                      三 跨月判据 = 年或月任一变化（同一月内不重复换表）；
                      四 负增量（表计回卷 / 换表）不计入并置信息级成因，不置故障；
                      五 无全局变量、无外部变量声明、无物理地址寻址。
  输出契约 Output contract:
                      eLevel 四级互斥；bWarn 在预警及以上为真，bOver 仅超限为真；
                      bMonthRoll 为跨月单拍脉冲（内部位置位、出口映射后撤销）；
                      非有限能耗增量不穿透出口（已用量保持上拍值）；
                      eCause 故障级成员均与 bError 配对（R45），信息级不置故障。
  修订记录 Revision  :
    2026-11-20  v1.0.0  R55 首版（批 1 · 序号 3）
  ==================================================================
*)

TYPE E_DL_EngLevel :
(
    eNormal := 0,       // 正常：占用低于预警阈 / normal, occupancy below the warning threshold
    eWarn   := 10,      // 预警：占用达预警阈 / warning, occupancy reached the warning threshold
    eCrit   := 20,      // 临界：占用达临界阈 / critical, occupancy reached the critical threshold
    eOver   := 30       // 超限：占用越过 100% / over, occupancy beyond one hundred percent
);
END_TYPE

TYPE E_DL_EngCause :
(
    eNone       := 0,   // 无成因 / no cause
    eCfgIllegal := 1,   // 组态非法：月/日/阈值或预算表越域（故障级）/ illegal config, month, day, threshold or budget table out of domain
    eBudgetZero := 2,   // 当月预算非正，占用率不可算（故障级）/ current month budget not positive, occupancy not computable
    eNegDelta   := 3,   // 负增量已忽略（信息级，不置故障）/ negative increment ignored, informational without a fault
    eBadDelta   := 4    // 增量非有限已忽略（信息级，不置故障）/ non-finite increment ignored, informational without a fault
);
END_TYPE

FUNCTION_BLOCK FB_DL_EnergyMonthPreset
VAR_INPUT
    bEnable          : BOOL := TRUE;         // 使能，下降沿冻结累计并按使能沿重建 / enable, falling edge freezes accumulation, the rising edge rebuilds it
    bReset           : BOOL := FALSE;         // 复位上升沿清当月累计与告警 [-] / reset rising edge clears the monthly accumulation and alarms
    nYear            : INT := 2026;           // 当前年份 [年]，域 2000..2100 / current year [year], domain 2000 to 2100
    nMonth           : INT := 1;              // 当前月份 [月]，域 1..12 / current month [month], domain 1 to 12
    nDayOfMonth      : INT := 1;              // 当月第几日 [日]，域 1..31 / day of month [day], domain 1 to 31
    bEnergyPulse     : BOOL := FALSE;         // 能耗增量脉冲，上升沿计入一次 [-] / energy increment pulse, counted once on the rising edge
    fEnergyDeltaKwh  : REAL := 0.0;           // 单次脉冲的能耗增量 [千瓦时] / energy increment per pulse [kilowatt hour]
    fBudgetOverrideKwh: REAL := 0.0;          // 预算覆盖值，大于零时取代预置表 [千瓦时] / budget override, replaces the table when positive [kilowatt hour]
    fWarnPct         : REAL := 90.0;          // 预警阈，占预算百分比 [百分比] / warning threshold as a percentage of the budget [percent]
    fCritPct         : REAL := 95.0;          // 临界阈，占预算百分比 [百分比] / critical threshold as a percentage of the budget [percent]
END_VAR
VAR_IN_OUT
    afMonthBudgetKwh : ARRAY[1..12] OF REAL;  // 12 个月预算预置表，下标即月份 [千瓦时]，引用型入参由调用方持有 / twelve month budget preset table, subscript is the month [kilowatt hour], reference parameter owned by the caller
END_VAR
VAR_OUTPUT
    fUsedKwh         : REAL := 0.0;           // 当月已用能耗 [千瓦时] / energy used in the current month [kilowatt hour]
    fBudgetKwh       : REAL := 0.0;           // 当月生效预算 [千瓦时] / effective budget of the current month [kilowatt hour]
    fRemainKwh       : REAL := 0.0;           // 当月剩余预算 [千瓦时]，可为负 / remaining budget of the current month, may be negative [kilowatt hour]
    fUsedPct         : REAL := 0.0;           // 当月预算占用百分比 [百分比] / monthly budget occupancy [percent]
    fDailyAvgKwh     : REAL := 0.0;           // 当月日均能耗 [千瓦时每日] / month to date daily average energy [kilowatt hour per day]
    fProjMonthKwh    : REAL := 0.0;           // 按日均推算的月末能耗 [千瓦时] / month end projection from the daily average [kilowatt hour]
    eLevel           : E_DL_EngLevel := E_DL_EngLevel.eNormal; // 预算级别出口 [枚举] / budget level outlet [enum]
    bWarn            : BOOL := FALSE;         // 预警及以上标志 [-] / warning and above flag
    bOver            : BOOL := FALSE;         // 超限标志 [-] / over budget flag
    bMonthRoll       : BOOL := FALSE;         // 跨月换表单拍脉冲 [-] / month rollover single-shot pulse
    nMonthActive     : INT := 0;              // 当前生效月份 [月] / currently active month [month]
    eCause           : E_DL_EngCause := E_DL_EngCause.eNone; // 成因出口 [枚举] / cause outlet [enum]
    bError           : BOOL := FALSE;         // 故障锁存标志 [-] / fault latch flag
END_VAR
VAR
    rtEnergy         : R_TRIG;                // 能耗脉冲沿检测，段 0 无条件刷新 / energy pulse edge detector, refreshed unconditionally in segment zero
    rtReset          : R_TRIG;                // 复位沿检测，段 0 无条件刷新 / reset edge detector, refreshed unconditionally in segment zero
    _eLevel          : E_DL_EngLevel := E_DL_EngLevel.eNormal;  // 内部级别，锁存至下拍重算 / internal level, recomputed every scan
    _eCause          : E_DL_EngCause := E_DL_EngCause.eNone;   // 内部信息级成因，每拍重算 / internal informational cause, recomputed every scan
    _eFaultCause     : E_DL_EngCause := E_DL_EngCause.eNone;   // 内部故障级成因，锁存至复位沿 / internal fault cause, latched until the reset edge
    _bFault          : BOOL := FALSE;         // 故障锁存位（组态类成因）/ fault latch bit for configuration causes
    _bMonthRollInt   : BOOL := FALSE;         // 跨月脉冲内部位，统一出口映射 / internal rollover pulse bit, mapped at the unified outlet
    _bInit           : BOOL := FALSE;         // 首扫初始化完成标志（R310）/ first scan initialisation flag
    _bMonthOk        : BOOL := FALSE;         // 年/月/日域闸通过 [-] / year, month and day domain gate passed
    _bDeltaUsable    : BOOL := FALSE;         // 本拍增量可计入 [-] / this scan increment is countable
    _bNegDelta       : BOOL := FALSE;         // 本拍增量为负 [-] / this scan increment is negative
    _bBadDelta       : BOOL := FALSE;         // 本拍增量非有限 [-] / this scan increment is non-finite
    _bDayOk          : BOOL := FALSE;         // 当日序号可用于日均分母 [-] / day index usable as the daily divisor
    _nYearPrev       : INT := 0;              // 上一拍年份快照 [年] / previous scan year snapshot [year]
    _nMonthPrev      : INT := -1;             // 上一拍月份快照，初值 -1 保证首拍必换表 [月] / previous scan month snapshot, minus one forces a rollover on the first scan
    _nMonthUse       : INT := 1;              // 钳定后的月份 [月] / clamped month [month]
    _nDayUse         : INT := 1;              // 钳定后的当日序号 [日] / clamped day index [day]
    _nDaysInMonth    : INT := 30;             // 当月日历天数 [日] / calendar days of the current month [day]
    _fBudgetUse      : REAL := 0.0;           // 生效预算暂存 [千瓦时] / effective budget held in a local [kilowatt hour]
    _fDeltaUse       : REAL := 0.0;           // 本拍计入的增量 [千瓦时] / increment actually counted this scan [kilowatt hour]
    _fUsed           : REAL := 0.0;           // 累计已用量保持块 [千瓦时] / accumulated energy holder [kilowatt hour]
    _fUsedAcc        : REAL := 0.0;           // 累计已用量工作值 [千瓦时] / accumulated energy working value [kilowatt hour]
    _fPct            : REAL := 0.0;           // 占用率工作值 [百分比] / occupancy working value [percent]
    _fRemain         : REAL := 0.0;           // 剩余量工作值 [千瓦时] / remaining working value [kilowatt hour]
    _fDaily          : REAL := 0.0;           // 日均工作值 [千瓦时每日] / daily average working value [kilowatt hour per day]
    _fProj           : REAL := 0.0;           // 月末预测工作值 [千瓦时] / projection working value [kilowatt hour]
    _fDayDiv         : REAL := 1.0;           // 日均除子（当日序号）[日] / daily divisor, the day index [day]
END_VAR
VAR CONSTANT
    DL_EMP_WARNPCT_MIN : REAL := 1.0;         // 预警阈下限 [百分比] / warning threshold floor [percent]
    DL_EMP_CRITPCT_MAX : REAL := 100.0;       // 临界阈上限 [百分比] / critical threshold ceiling [percent]
    DL_EMP_USED_MAX    : REAL := 1.0E12;      // 已用量上限，防累计溢出失真 [千瓦时] / used energy ceiling against accumulation distortion [kilowatt hour]
    DL_EMP_DELTA_MAX   : REAL := 1.0E7;       // 单次增量上限，防量纲错配放大 [千瓦时] / single increment ceiling against a dimension mismatch [kilowatt hour]
    DL_EMP_DAY_MAX     : INT := 31;           // 月内最大天数 [日] / maximum days within a month [day]
    DL_EMP_YEAR_MIN    : INT := 2000;         // 年份下限 [年] / year floor [year]
    DL_EMP_YEAR_MAX    : INT := 2100;         // 年份上限 [年] / year ceiling [year]
END_VAR

// 段 0｜沿检测无条件周期刷新（禁入分支）/ segment 0, unconditional refresh of the edge detectors, never inside a branch
rtEnergy(CLK := bEnergyPulse); // 能耗脉冲沿无条件刷新 / unconditional refresh of the energy pulse edge
rtReset(CLK := bReset); // 复位沿无条件刷新 / unconditional refresh of the reset edge

// 段 1｜首扫初始化（R310）：月份快照置 -1 使首拍必走一次换表 / segment 1, first scan initialisation, the month snapshot at minus one forces one rollover on the first scan
IF NOT _bInit THEN // 首扫一拍 / the very first scan
    _bInit := TRUE; // 置首扫完成标志 / raise the first scan flag
    _nMonthPrev := -1; // 月份快照置非法值 / put the month snapshot at an illegal value
    _nYearPrev := 0; // 年份快照清零 / clear the year snapshot
    _fUsed := 0.0; // 已用量清零 / clear the accumulated energy
    _bFault := FALSE; // 故障锁存清零 / clear the fault latch
    _eCause := E_DL_EngCause.eNone; // 信息级成因清零 / clear the informational cause
    _eFaultCause := E_DL_EngCause.eNone; // 故障级成因清零 / clear the fault cause
END_IF

// 段 2｜域闸：年月日、阈值对、预置表逐项（R151 全覆盖）/ segment 2, domain gate over year, month, day, the threshold pair and the preset table
_bMonthOk := TRUE; // 域闸标志预置通过 / preset the domain gate flag to passed
IF (nYear < DL_EMP_YEAR_MIN) OR (nYear > DL_EMP_YEAR_MAX) THEN // 年份越域 / year out of domain
    _bMonthOk := FALSE; // 判越域 / mark out of domain
END_IF
IF (nMonth < 1) OR (nMonth > 12) THEN // 月份越域 / month out of domain
    _bMonthOk := FALSE; // 判越域 / mark out of domain
END_IF
IF (nDayOfMonth < 1) OR (nDayOfMonth > DL_EMP_DAY_MAX) THEN // 当日序号越域 / day index out of domain
    _bMonthOk := FALSE; // 判越域 / mark out of domain
END_IF
IF (fWarnPct < DL_EMP_WARNPCT_MIN) OR (fWarnPct > DL_EMP_CRITPCT_MAX) OR (fWarnPct <> fWarnPct) THEN // 预警阈越域或非有限 / warning threshold out of domain or non-finite
    _bMonthOk := FALSE; // 判越域 / mark out of domain
END_IF
IF (fCritPct < fWarnPct) OR (fCritPct > DL_EMP_CRITPCT_MAX) OR (fCritPct <> fCritPct) THEN // 临界阈低于预警阈或越域 / critical threshold below the warning threshold or out of domain
    _bMonthOk := FALSE; // 判越域 / mark out of domain
END_IF
IF (fBudgetOverrideKwh <> fBudgetOverrideKwh) OR (fBudgetOverrideKwh < 0.0) THEN // 预算覆盖值非有限或为负 / budget override non-finite or negative
    _bMonthOk := FALSE; // 判越域 / mark out of domain
END_IF
IF _bMonthOk THEN // 域内才可安全读预置表 / the preset table is only read inside the domain
    _nMonthUse := nMonth; // 月份直通 / month passes through
    _nDayUse := nDayOfMonth; // 当日序号直通 / day index passes through
ELSE // 域外走两级回退（R117）/ out of domain uses the two stage fallback
    _nMonthUse := 1; // 一级：月份回默认一 / stage one, the month falls back to one
    _nDayUse := 1; // 一级：当日回默认一 / stage one, the day falls back to one
    IF NOT _bFault THEN // 未锁存才记故障 / record the fault only when not yet latched
        _eFaultCause := E_DL_EngCause.eCfgIllegal; // 故障级成因记组态非法 / record the illegal configuration cause
        _bFault := TRUE; // 置故障锁存 / raise the fault latch
    END_IF
END_IF

// 段 3｜换表判据：年或月任一变化即换表，首拍必换；同年同月不重复换表 / segment 3, rollover when the year or the month changed, mandatory on the first scan
IF (_nMonthUse <> _nMonthPrev) OR (nYear <> _nYearPrev) THEN // 跨月或跨年 / month or year changed
    _nMonthPrev := _nMonthUse; // 月份快照推进 / advance the month snapshot
    _nYearPrev := nYear; // 年份快照推进 / advance the year snapshot
    _fUsed := 0.0; // 换表清零当月累计 / clear the monthly accumulation on rollover
    _bMonthRollInt := TRUE; // 跨月脉冲内部位置位（出口映射后撤销）/ raise the internal rollover bit, revoked after outlet mapping
    _eCause := E_DL_EngCause.eNone; // 换表清信息级成因（跨月是正常事件）/ clear the informational cause, a rollover is a normal event
END_IF

// 段 4｜预算取值：覆盖值优先，其次预置表；两项都非正判故障 / segment 4, effective budget, the override first and the preset table second, both non-positive is a fault
_fBudgetUse := 0.0; // 生效预算预置零 / preset the effective budget to zero
IF fBudgetOverrideKwh > 0.0 THEN // 覆盖值生效 / the override is effective
    _fBudgetUse := fBudgetOverrideKwh; // 取覆盖值 / take the override
ELSE // 覆盖值未给 / the override is absent
    _fBudgetUse := afMonthBudgetKwh[_nMonthUse]; // 按钳定月份取预置值，下标 1..12 已回钳 / read the preset by the clamped month, the index is already inside one through twelve
END_IF
IF (_fBudgetUse <> _fBudgetUse) OR ((_fBudgetUse - _fBudgetUse) <> (_fBudgetUse - _fBudgetUse)) THEN // 预算非有限 / budget non-finite
    _fBudgetUse := 0.0; // 非有限归零，绝不进除法 / zeroed so nothing non-finite enters a division
END_IF
IF _fBudgetUse <= 0.0 THEN // 预算非正 / budget not positive
    IF NOT _bFault THEN // 未锁存才记故障 / record the fault only when not yet latched
        _eFaultCause := E_DL_EngCause.eBudgetZero; // 故障级成因记预算非正 / record the non-positive budget cause
        _bFault := TRUE; // 置故障锁存 / raise the fault latch
    END_IF
END_IF

// 段 5｜增量计入：仅上升沿、仅有限、仅非负；负与非有限各记信息级成因 / segment 5, increment only on the rising edge, only finite, only non-negative
_bDeltaUsable := FALSE; // 可计入标志预置假 / preset the countable flag to false
_bNegDelta := FALSE; // 负增量标志预置假 / preset the negative increment flag to false
_bBadDelta := FALSE; // 非有限增量标志预置假 / preset the non-finite increment flag to false
_fDeltaUse := 0.0; // 本拍计入量预置零 / preset the counted increment to zero
IF rtEnergy.Q THEN // 脉冲上升沿 / rising edge of the pulse
    IF (fEnergyDeltaKwh <> fEnergyDeltaKwh) OR ((fEnergyDeltaKwh - fEnergyDeltaKwh) <> (fEnergyDeltaKwh - fEnergyDeltaKwh)) THEN // 增量非有限 / increment non-finite
        _bBadDelta := TRUE; // 置非有限标志 / raise the non-finite flag
    ELSIF fEnergyDeltaKwh < 0.0 THEN // 增量为负（表计回卷或换表）/ increment negative, meter rollback or replacement
        _bNegDelta := TRUE; // 置负增量标志 / raise the negative flag
    ELSIF fEnergyDeltaKwh > DL_EMP_DELTA_MAX THEN // 增量越上限 / increment above the ceiling
        _fDeltaUse := DL_EMP_DELTA_MAX; // 上钳，防量纲错配放大 / clamp upward against a dimension mismatch
        _bDeltaUsable := TRUE; // 置可计入标志 / raise the countable flag
    ELSE // 正常增量 / normal increment
        _fDeltaUse := fEnergyDeltaKwh; // 直通计入 / counted as received
        _bDeltaUsable := TRUE; // 置可计入标志 / raise the countable flag
    END_IF
END_IF
_eCause := E_DL_EngCause.eNone; // 信息级成因每拍重算 / the informational cause is recomputed every scan
IF _bNegDelta THEN // 负增量拍 / negative increment scan
    _eCause := E_DL_EngCause.eNegDelta; // 信息级成因，不置故障（R45 反向：信息级不配对 bError）/ informational cause without a fault
ELSIF _bBadDelta THEN // 非有限增量拍 / non-finite increment scan
    _eCause := E_DL_EngCause.eBadDelta; // 信息级成因，不置故障 / informational cause without a fault
END_IF

// 段 6｜累计与复位：复位沿清当月累计；累计上限饱和并置信息级成因 / segment 6, accumulation and reset, with saturation at the ceiling
_fUsedAcc := _fUsed; // 工作值取保持值 / the working value takes the holder
IF rtReset.Q THEN // 复位沿 / reset edge
    _fUsedAcc := 0.0; // 当月累计清零 / clear the monthly accumulation
END_IF
IF _bDeltaUsable THEN // 本拍有可计入增量 / a countable increment exists this scan
    _fUsedAcc := _fUsedAcc + _fDeltaUse; // 累加 / accumulate
    IF _fUsedAcc > DL_EMP_USED_MAX THEN // 累计越上限 / accumulation above the ceiling
        _fUsedAcc := DL_EMP_USED_MAX; // 饱和到上限 / saturate at the ceiling
    END_IF
END_IF
IF NOT bEnable THEN // 失能：冻结保持末值（R191 显式声明）/ disabled, freeze and hold the last value as declared
    _fUsedAcc := _fUsed; // 冻结保持，不再累加 / freeze and hold without further accumulation
END_IF
_fUsed := _fUsedAcc; // 保持块更新 / refresh the holder

// 段 7｜日历天数与日均：闰年二月按 29 日；除子先域闸 / segment 7, calendar days and daily average, the divisor is gated first
_nDaysInMonth := 31; // 默认 31 日 / default thirty one days
CASE _nMonthUse OF
1, 3, 5, 7, 8, 10, 12: // 大月 / long months
    _nDaysInMonth := 31; // 三十一日 / thirty one days
2: // 二月 / february
    IF ((nYear MOD 4) = 0) AND (((nYear MOD 100) <> 0) OR ((nYear MOD 400) = 0)) THEN // 闰年判据 / leap year criterion
        _nDaysInMonth := 29; // 闰年二月二十九日 / twenty nine days in a leap year
    ELSE
        _nDaysInMonth := 28; // 平年二月二十八日 / twenty eight days in a common year
    END_IF
4, 6, 9, 11: // 小月 / short months
    _nDaysInMonth := 30; // 三十日 / thirty days
ELSE // 非法月份兜底（R128）/ illegal month fallback
    _nDaysInMonth := 30; // 兜底三十日 / fall back to thirty days
END_CASE
_bDayOk := (_nDayUse >= 1) AND (_nDayUse <= _nDaysInMonth); // 当日序号在日历域内 / the day index is inside the calendar domain
IF _bDayOk THEN // 除子可用 / the divisor is usable
    _fDayDiv := _nDayUse; // 除子取当日序号，已证 不小于 1 / the divisor takes the day index, proven not below one
ELSE
    _fDayDiv := 1.0; // 回退为 1，防除零 / fall back to one against division by zero
END_IF

// 段 8｜占用率与分级：预算非正时不计算占用率，级别保持上拍 / segment 8, occupancy and grading, skipped when the budget is not positive
IF _fBudgetUse > 0.0 THEN // 预算可用 / the budget is usable
    _fPct := _fUsed / _fBudgetUse * 100.0; // 占用率，除子已证大于零 / occupancy, divisor proven positive
    _fRemain := _fBudgetUse - _fUsed; // 剩余量（可为负）/ remaining budget, may be negative
    _fDaily := _fUsed / _fDayDiv; // 日均能耗，除子已证不小于 1 / daily average, divisor proven not below one
    _fProj := _fDaily * INT_TO_REAL(_nDaysInMonth); // 月末预测，乘数为日历天数 / month end projection over the calendar days
    IF _fPct >= 100.0 THEN // 越过全额 / beyond the full budget
        _eLevel := E_DL_EngLevel.eOver; // 超限级 / over level
    ELSIF _fPct >= fCritPct THEN // 达临界阈 / reached the critical threshold
        _eLevel := E_DL_EngLevel.eCrit; // 临界级 / critical level
    ELSIF _fPct >= fWarnPct THEN // 达预警阈 / reached the warning threshold
        _eLevel := E_DL_EngLevel.eWarn; // 预警级 / warning level
    ELSE
        _eLevel := E_DL_EngLevel.eNormal; // 正常级 / normal level
    END_IF
END_IF

// 段 9｜统一出口：脉冲映射、名实双出口、故障与级别落定 / segment 9, unified outlet for the pulse, the matched flags and the level
bMonthRoll := _bMonthRollInt; // 跨月脉冲映射本拍值 / map the rollover pulse for this scan
_bMonthRollInt := FALSE; // 映射后立即撤销，保证单拍宽度（R187 两段式）/ revoke right after mapping to keep a single-scan width
fUsedKwh := _fUsed; // 已用量出口 / used energy outlet
fBudgetKwh := _fBudgetUse; // 生效预算出口 / effective budget outlet
fRemainKwh := _fRemain; // 剩余量出口 / remaining budget outlet
fUsedPct := _fPct; // 占用率出口 / occupancy outlet
fDailyAvgKwh := _fDaily; // 日均出口 / daily average outlet
fProjMonthKwh := _fProj; // 月末预测出口 / projection outlet
eLevel := _eLevel; // 级别出口单点映射 / single-point level outlet mapping
bWarn := (_eLevel = E_DL_EngLevel.eWarn) OR (_eLevel = E_DL_EngLevel.eCrit) OR (_eLevel = E_DL_EngLevel.eOver); // 预警及以上（挂状态量）/ warning and above, a state quantity
bOver := (_eLevel = E_DL_EngLevel.eOver); // 超限（挂状态量）/ over budget, a state quantity
nMonthActive := _nMonthUse; // 生效月份出口 / active month outlet
IF _bFault THEN // 故障锁存优先 / the fault latch takes priority
    eCause := _eFaultCause; // 故障级成因锁存回放（禁按当下输入重推断）/ the fault cause is replayed from the latch
ELSE
    eCause := _eCause; // 信息级成因直映 / the informational cause is mapped directly
END_IF
bError := _bFault; // 故障标志与锁存位同源 / the fault flag shares the latch source
END_FUNCTION_BLOCK

(* ---- FB_DL_EnthalpyChangeover.st ---- *)
(*==============================================================================
 * 组件名称 (Component)  : FB_DL_EnthalpyChangeover
 * 所属子库 (Sublibrary) : DL_Process
 * 前缀     (Prefix)     : FB_DL_
 * 当前版本 (Version)    : 1.0.0
 * 兼容性   (Platform)   : CODESYS 3.5 / TwinCAT 3 / 汇川 InoProShop / Schneider
 *                         Machine Expert；纯 IEC 61131-3（第 3 版），
 *                         仅依赖标准库 TON，零厂商方言
 * 作者     (Author)     : 道莅代码库 · PLC编程专家（R31）
 * 开源溯源 (Origin)     : 空调系统新风/回风焓值优先切换公开控制语义
 *                         （T1-2 ROOM_CONTROL 族行为定义），道莅 clean-room
 *                         防御性实现，未复制任何外部源码行
 * 功能描述 (Function)   : 新风/回风焓值优先模式仲裁件（模式仲裁层）。自动态以
 *                         「新风焓 < 回风焓 − 死区」判新风优先，带回差不对称
 *                         双向判定防振荡；手动态直通锁存；每次切换经最小驻留
 *                         时间抑制频切。与已收口 FB_DL_EnthalpyCompareCtrl
 *                         （单回路执行块）的职责边界：本件只决定用哪路风源，
 *                         不执行风阀/风机动作。
 * 码位     (Codes)      : 16#0005_008F 信息级：焓值非有限保持上次选择、
 *                         fDiffMin 负值钳 0、驻留期切换请求被拒（不置 bError）
 *                         16#0005_0090~0093 故障级保留未启用（本轮无故障级条件，
 *                         码表与实现对齐，不虚声明）
 * 边界防错 (Boundary)   : 1 任一焓值非有限（x<>x 自反判加幅值界）保持上次选择；
 *                         2 fDiffMin<0 钳 0 记信息码；3 首拍初始化为回风（保守侧）；
 *                         4 TON 每拍无条件刷新，驻留重置经单拍断输入实现；
 *                         5 非法枚举走 CASE ELSE 保持现状记信息码。
 * 修订历史 (Revision)   : 2026-11-18 v1.0.0 首版入库（R31 · 阶段三 · 序 3）
 *==============================================================================*)

(*------------------------------------------------------------------------------
 * 枚举: E_DL_ChangeoverMode（归属本功能块，同文件发布，全库唯一属主）
 *----------------------------------------------------------------------------*)
TYPE E_DL_ChangeoverMode :
(
    eAuto      := 0,    // 自动态：按焓差判据仲裁 / Auto, arbitrate by enthalpy difference
    eManualOA  := 10,   // 手动新风：直通锁存新风侧 / Manual fresh air, direct select
    eManualRA  := 20    // 手动回风：直通锁存回风侧 / Manual return air, direct select
);
END_TYPE

(*------------------------------------------------------------------------------
 * 枚举: E_DL_AirSource（归属本功能块，同文件发布，全库唯一属主）
 *----------------------------------------------------------------------------*)
TYPE E_DL_AirSource :
(
    eOA := 0,         // 新风源 / Outside air source
    eRA := 10         // 回风源 / Return air source
);
END_TYPE

(*==============================================================================
 * 功能块: FB_DL_EnthalpyChangeover
 * 调用约定: 每个扫描周期无条件调用一次；焓值由调用方用 FC_DL_HumidAirEnthalpy
 *           预算后经引脚注入，本件不做焓值计算。
 *==============================================================================*)
FUNCTION_BLOCK FB_DL_EnthalpyChangeover
VAR_INPUT
    fEnthOA    : REAL := 0.0;          // 新风焓值 [kJ/kg]，调用方预算注入 / Outside air enthalpy [kJ/kg]
    fEnthRA    : REAL := 0.0;          // 回风焓值 [kJ/kg]，调用方预算注入 / Return air enthalpy [kJ/kg]
    fDiffMin   : REAL := 2.0;          // 新风优先判据死区 [kJ/kg]，负值钳 0 / Minimum benefit deadband [kJ/kg]
    tMinDwell  : TIME := T#120S;       // 切换最小驻留 [ms]，抑制频切 / Minimum dwell time [ms] against hunting
    eMode      : E_DL_ChangeoverMode;  // 运行模式选择 / Operating mode selector
    bEn        : BOOL := FALSE;        // 使能 / Enable flag
END_VAR
VAR_OUTPUT
    eSelect    : E_DL_AirSource;       // 当前风源选择 / Selected air source
    bSwitching : BOOL;                 // 切换进行中单拍脉冲 / Switching pulse, one scan per change
    uErrorId   : UDINT;                // 信息级码，0 = 无信息 / Info code, 0 = none
END_VAR
VAR
    tonDwell   : TON;                  // 最小驻留定时器，每拍无条件刷新 / Dwell timer, refreshed every scan
    bFirstScan : BOOL := TRUE;         // 首扫初始化标志 / First-scan initialisation flag
    bDwellRst  : BOOL;                 // 本拍驻留重置请求（单拍断输入）/ One-scan dwell reset request
    bWantOA    : BOOL;                 // 本拍新风侧请求 / Fresh air request this scan
    bWantRA    : BOOL;                 // 本拍回风侧请求 / Return air request this scan
    bGrant     : BOOL;                 // 本拍请求获准切换 / Request granted this scan
    bFinite    : BOOL;                 // 焓值双端有限标志 / Both enthalpies finite flag
    fDiffEff   : REAL;                 // 钳位后生效死区 [kJ/kg] / Effective clamped deadband [kJ/kg]
    fMargin    : REAL;                 // 回风减新风焓差 [kJ/kg] / Enthalpy margin RA minus OA [kJ/kg]
    bParamClamp: BOOL;                 // 参数钳位信息标志 / Parameter clamp info flag
END_VAR
VAR CONSTANT
    DL_ECO_FIN    : REAL := 1.0E30;    // REAL 有限幅值判界 / REAL finiteness magnitude bound
    DL_ECO_BACK   : REAL := 0.5;       // 不对称回差系数：回切阈 = 死区乘该系数 / Asymmetric hysteresis factor for switching back
END_VAR

// ---- 段 1｜定时器无条件刷新（红线：禁入条件分支）------------------------------
tonDwell(IN := (NOT bDwellRst), PT := tMinDwell);     // 驻留计时，重置拍断输入 / Dwell timing, broken input on reset scan

// ---- 段 2｜首拍初始化为回风（保守侧）------------------------------------------
IF bFirstScan THEN
    eSelect    := eRA;                                // 首拍保守选回风 / Conservative return air on first scan
    bFirstScan := FALSE;                              // 清首扫标志 / Clear first-scan flag
END_IF

// ---- 段 3｜参数与输入有效性 ----------------------------------------------------
bParamClamp := FALSE;                                 // 钳位信息先清 / Clear clamp info
fDiffEff := fDiffMin;                                 // 死区原值 / Deadband as-is
IF fDiffEff < 0.0 THEN
    fDiffEff := 0.0;                                  // 负死区钳 0 / Clamp negative deadband to zero
    bParamClamp := TRUE;                              // 记参数钳位 / Record parameter clamp
END_IF
bFinite := (fEnthOA = fEnthOA) AND (fEnthRA = fEnthRA)
       AND (ABS(fEnthOA) < DL_ECO_FIN) AND (ABS(fEnthRA) < DL_ECO_FIN); // 焓值双端有限 / Both enthalpies finite

// ---- 段 4｜请求生成（非有限与非法模式一律保持现状 + 信息码）--------------------
bWantOA := FALSE;                                     // 请求先清 / Clear requests
bWantRA := FALSE;                                     // 请求先清 / Clear requests
IF NOT bFinite THEN
    uErrorId := 16#0005_008F;                         // 信息级：焓值非有限保持现状 / Info: non-finite, hold selection
ELSIF eMode = eAuto THEN
    fMargin := fEnthRA - fEnthOA;                     // 回风减新风焓差 / Enthalpy margin
    IF (eSelect = eRA) AND (fMargin > fDiffEff) THEN
        bWantOA := TRUE;                              // 进新风：收益须超死区（正向全阈）/ Enter OA only above full deadband
    ELSIF (eSelect = eOA) AND (fMargin < fDiffEff * DL_ECO_BACK) THEN
        bWantRA := TRUE;                              // 退回风：低于半阈即回（不对称回差）/ Back to RA below half threshold
    END_IF
    uErrorId := 16#0000_0000;                         // 自动态正常清码 / Clear code in normal auto
ELSIF eMode = eManualOA THEN
    bWantOA := TRUE;                                  // 手动新风直通 / Manual OA direct
    uErrorId := 16#0000_0000;                         // 手动正常清码 / Clear code in manual
ELSIF eMode = eManualRA THEN
    bWantRA := TRUE;                                  // 手动回风直通 / Manual RA direct
    uErrorId := 16#0000_0000;                         // 手动正常清码 / Clear code in manual
ELSE
    uErrorId := 16#0005_008F;                         // 非法模式兜底保持现状 / Illegal mode fallback, hold
END_IF
IF bParamClamp AND (uErrorId = 16#0000_0000) THEN
    uErrorId := 16#0005_008F;                         // 钳位信息并码（信息级槽合并复用）/ Merge clamp info into info slot
END_IF

// ---- 段 5｜驻留门控与切换执行 --------------------------------------------------
bGrant := FALSE;                                      // 获准标志先清 / Clear grant flag
IF bEn AND (bWantOA <> bWantRA) AND (tonDwell.Q) THEN
    IF bWantOA AND (eSelect = eRA) THEN
        eSelect    := eOA;                            // 切到新风 / Switch to outside air
        bGrant     := TRUE;                           // 本拍获准 / Granted this scan
    ELSIF bWantRA AND (eSelect = eOA) THEN
        eSelect    := eRA;                            // 切到回风 / Switch to return air
        bGrant     := TRUE;                           // 本拍获准 / Granted this scan
    END_IF
ELSIF bEn AND (bWantOA <> bWantRA) AND (NOT tonDwell.Q) THEN
    uErrorId := 16#0005_008F;                         // 信息级：驻留期切换请求被拒 / Info: request rejected in dwell
END_IF
bSwitching := bGrant;                                 // 切换脉冲单拍有效 / One-scan switching pulse
bDwellRst  := bGrant;                                 // 获准拍断驻留输入重置计时 / Break dwell input on granted scan

// ---- 段 6｜非使能保持：不改变选择，仅清切换脉冲 --------------------------------
IF NOT bEn THEN
    bSwitching := FALSE;                              // 非使能清脉冲 / Clear pulse when disabled
END_IF
END_FUNCTION_BLOCK

(* ---- FB_DL_EnthalpyPrioritySwitch.st ---- *)
(*
  Name        : FB_DL_EnthalpyPrioritySwitch
  Category    : DL_Process
  Version     : 1.0.0
  Purpose     : 焓值优先切换：新风/回风焓差判据经迟滞双阈 + 驻留确认切换经济器模式，出口为模式枚举（与焓差判定件职责分立）；/ Enthalpy priority switch: outside/return air enthalpy difference through hysteresis band with dwell confirmation switches economizer mode, mode-enum outlet only
  溯源        : 借 oscat-building 的焓值优先切换待挖组织，clean-room 实现
  Boundary    : ① 焓差迟滞带双阈组态闸：切换阈 > 返回阈否则锁存故障（相等不立）；
                ② 切换判据须持续 tHold 驻留才生效（防高频抖动），驻留 TON 断输入归零（R40）；
                ③ 任一温度/湿度派生焓值非有限 → 保持当前模式 + bSensorBad 当拍出口（不切到未知工况）；
                ④ 最小驻留双侧对称：新模式下判据同样须持续 tHold 才切回（双向同参数天然对称）；
                ⑤ 与 R6 焓差判据件分工：本件只输出模式枚举，不做焓差报警（职责不重叠）；
                ⑥ 焓值由属主计算输入，本件零焓值公式内嵌（单一职责）。
*)
TYPE E_DL_EntMode :
(
    eRecirc := 0,                            (* 回风循环模式（经济器关闭） / Recirculation mode *)
    eEcon   := 10                            (* 经济器模式（新风优先） / Economizer mode *)
);
END_TYPE

TYPE E_DL_EntState :
(
    eIdle  := 0,                             (* 未使能（模式保持） / Disabled, mode held *)
    eRun   := 10,                            (* 切换仲裁运行 / Arbitration running *)
    eFault := 90                             (* 故障锁存相 / Fault latched *)
);
END_TYPE

TYPE E_DL_EntCause :
(
    eNone      := 0,                         (* 无成因 / No cause *)
    eCfgIllegal:= 1,                        (* 组态非法：迟滞带倒挂/驻留越域 / Illegal config *)
    ePhaseBad  := 2                         (* 非法相位兜底 / Illegal phase fallback *)
);
END_TYPE

FUNCTION_BLOCK FB_DL_EnthalpyPrioritySwitch
VAR_INPUT
    fHOut    : REAL := 30.0;                 (* 新风焓值（属主计算输入）[kJ/kg] / Outside air enthalpy *)
    fHRet    : REAL := 40.0;                 (* 回风焓值（属主计算输入）[kJ/kg] / Return air enthalpy *)
    fSwOn    : REAL := 2.0;                  (* 切换阈：焓差超过此值切经济器，域 > 返回阈 [kJ/kg] / Switch-on threshold *)
    fSwOff   : REAL := 0.5;                  (* 返回阈：焓差低于此值切回循环 [kJ/kg] / Switch-back threshold *)
    tHold    : TIME := T#120S;               (* 判据驻留时间，域 > T#0S [ms] / Dwell time *)
    tScan    : TIME := T#1S;                 (* 扫描周期，域 > T#0S [ms] / Scan period *)
    bEnable  : BOOL := TRUE;                 (* 使能 [-] / Enable *)
    bReset   : BOOL := FALSE;                (* 复位命令，上升沿清故障回循环模式 [-] / Reset command *)
END_VAR
VAR_OUTPUT
    eMode    : E_DL_EntMode;                 (* 当前模式出口（枚举，边界⑤） / Mode outlet *)
    bSensorBad: BOOL;                        (* 焓值失效当拍出口（边界③）[-] / Sensor bad outlet *)
    bEconAct : BOOL;                         (* 经济器激活指示（名实双出口）[-] / Economizer active indicator *)
    eState   : E_DL_EntState;                (* 状态出口 / State outlet *)
    eCause   : E_DL_EntCause;                (* 成因出口（R190 归因唯一） / Cause outlet *)
    bError   : BOOL;                         (* 故障锁存标志 [-] / Fault latch flag *)
END_VAR
VAR
    _eState : E_DL_EntState := E_DL_EntState.eIdle;  (* 内部相位（CASE 唯一写入目标） / Internal phase *)
    _eCause : E_DL_EntCause := E_DL_EntCause.eNone;  (* 成因锁存量 / Latched cause *)
    _eModeI : E_DL_EntMode := E_DL_EntMode.eRecirc;  (* 内部模式（初值循环侧，安全默认） / Internal mode *)
    rtReset : R_TRIG;                        (* 复位沿实例，段 0 无条件调用 / Reset edge instance *)
    tonHold : TON;                           (* 判据驻留计时（IN 串判据 + 相位闸，边界②④） / Dwell timer *)
    _bFault : BOOL;                          (* 故障锁存位 / Latched fault bit *)
    _bCfgBad: BOOL;                          (* 组态非法当拍量 / Illegal config this scan *)
    _bFinH  : BOOL;                          (* 双焓值有限性当拍量（边界③） / Enthalpies finiteness *)
    _bToEcon: BOOL;                          (* 切经济器判据当拍量 / To-economizer verdict *)
    _bToRec : BOOL;                          (* 切回循环判据当拍量 / To-recirc verdict *)
    _fDH    : REAL;                          (* 焓差中间量（回风 - 新风）[kJ/kg] / Enthalpy difference *)
END_VAR
VAR CONSTANT
    DL_ENT_EPS : REAL := 1.0E-6;             (* 判零容差 [-] / Epsilon *)
END_VAR

(* —— 段 0：当拍判据派生 + 实例无条件刷新（R228A；TON 段 0 无 IF 包裹，边界②） —— *)
_bCfgBad := NOT (fSwOn > fSwOff)                         (* 迟滞带组态闸：切换阈 > 返回阈（边界①） / Band config gate *)
            OR (fSwOff < (-DL_ENT_EPS))                  (* 返回阈非负域闸 / Return threshold gate *)
            OR NOT (tHold > T#0S) OR NOT (tScan > T#0S); (* 驻留/周期域闸（边界②） / Dwell and period gates *)
rtReset(CLK := bReset);                                  (* 复位沿每拍必调 / Reset edge every scan *)
_bFinH := (fHOut = fHOut) AND ((fHOut - fHOut) = (fHOut - fHOut))        (* 新风焓 NaN 自反 + Inf 差判闸（边界③） / Outdoor NaN and Inf gate *)
         AND (fHRet = fHRet) AND ((fHRet - fHRet) = (fHRet - fHRet));   (* 回风焓 NaN 自反 + Inf 差判闸 / Return NaN and Inf gate *)
_fDH := fHRet - fHOut;                                   (* 焓差 = 回风 - 新风（有限派生） / Enthalpy difference *)
IF NOT _bFinH THEN
    _fDH := 0.0;                                         (* 非有限拍焓差归零（判据失效不误切，边界③） / Difference zeroed *)
END_IF
_bToEcon := _bFinH AND (_fDH > fSwOn);                   (* 切经济器判据（迟滞上阈直比） / To-econ verdict *)
_bToRec := _bFinH AND (_fDH < fSwOff);                   (* 切回循环判据（迟滞下阈直比，边界②） / To-recirc verdict *)
tonHold(IN := ((_eState = E_DL_EntState.eRun) AND (_eModeI = E_DL_EntMode.eRecirc) AND _bToEcon)
             OR ((_eState = E_DL_EntState.eRun) AND (_eModeI = E_DL_EntMode.eEcon) AND _bToRec), PT := tHold);   (* 双向对称驻留（边界②④，R40） / Symmetric dwell timer *)

(* —— 段 1：单拍量预清零（R107） —— *)
bSensorBad := FALSE;                                     (* 传感器失效当拍出口预清 / Sensor bad preset *)
bEconAct := FALSE;                                       (* 激活指示出口预清（派生拍覆盖） / Active preset *)

(* —— 段 2：复位沿处理（作用域：清故障 + 模式回循环侧 + 迁 eIdle，R283 逐项声明） —— *)
IF rtReset.Q THEN
    _bFault := FALSE;                                    (* 清故障锁存 / Clear fault *)
    _eCause := E_DL_EntCause.eNone;                      (* 清成因 / Clear cause *)
    _eModeI := E_DL_EntMode.eRecirc;                     (* 模式回循环侧（安全默认） / Mode to recirculation *)
    eMode := E_DL_EntMode.eRecirc;                       (* 模式出口同步 / Mode outlet sync *)
    _eState := E_DL_EntState.eIdle;                      (* 迁未使能相 / Back to idle *)
END_IF

(* —— 段 3：组态故障锁存（锁存至复位沿，R189） —— *)
IF _bCfgBad AND NOT _bFault THEN
    _bFault := TRUE;                                     (* 锁存故障位 / Latch fault *)
    _eCause := E_DL_EntCause.eCfgIllegal;                (* 成因：组态非法 / Cause illegal config *)
    _eState := E_DL_EntState.eFault;                     (* 同步迁故障相 / Migrate to fault *)
END_IF

(* —— 段 4：CASE 主状态机（ELSE 兜底迁 eFault，红线 6） —— *)
CASE _eState OF
    E_DL_EntState.eIdle:                                 (* 未使能：模式出口保持确定值（状态镜像） / Idle *)
        eMode := _eModeI;                                (* 模式出口镜像（不留陈旧） / Mode outlet mirror *)
        IF bEnable AND NOT _bFault THEN
            _eState := E_DL_EntState.eRun;               (* 进入仲裁相 / Enter arbitration *)
        END_IF
    E_DL_EntState.eRun:                                  (* 仲裁相：判据 + 驻留 + 切换 / Arbitration *)
        IF NOT bEnable THEN
            _eState := E_DL_EntState.eIdle;              (* 失能回未使能（模式保持） / Back to idle *)
        ELSE
            IF NOT _bFinH THEN
                bSensorBad := TRUE;                      (* 焓值失效：保持当前模式（边界③） / Sensor bad hold *)
            ELSIF tonHold.Q THEN                         (* 判据持续满驻留：切换（边界②④） / Dwell elapsed, switch *)
                IF _eModeI = E_DL_EntMode.eRecirc THEN
                    _eModeI := E_DL_EntMode.eEcon;       (* 循环 → 经济器 / To economizer *)
                ELSE
                    _eModeI := E_DL_EntMode.eRecirc;     (* 经济器 → 循环（双向对称，边界④） / To recirculation *)
                END_IF
            END_IF
            eMode := _eModeI;                            (* 模式出口镜像（状态镜像，R191） / Mode outlet mirror *)
        END_IF
    E_DL_EntState.eFault:                                (* 故障相：模式冻结保持，仅复位沿出 / Fault *)
        eMode := _eModeI;                                (* 故障相模式出口保持镜像（确定值） / Mode mirror in fault *)
        ;                                                (* 锁存回放（R28） / Replay from latch *)
    ELSE                                                 (* 非法相位兜底迁安全态 / Illegal phase fallback *)
        _eState := E_DL_EntState.eFault; _bFault := TRUE;    (* 迁故障相 + 同步锁存 / To fault and latch *)
        _eCause := E_DL_EntCause.ePhaseBad;              (* 成因：非法相位 / Cause illegal phase *)
END_CASE

(* —— 段 5：出口映射（名实双出口，R191；bError/eState 同源） —— *)
bEconAct := (_eModeI = E_DL_EntMode.eEcon);              (* 经济器激活指示镜像 / Economizer active mirror *)
bError := _bFault;                                       (* 故障标志镜像 / Fault flag mirror *)
eState := _eState;                                       (* 状态出口 / State outlet *)
eCause := _eCause;                                       (* 成因出口 / Cause outlet *)
END_FUNCTION_BLOCK
